(* IEC 61131-3 sources: 2026_Projet_YGO_ExcavatriceDragage/CODE_BACKUP/CODE_20260902_JoyAvantHoming_v0.6.27/G_CYCLE, 4 files *)

(* ---- FB_Cycle.st ---- *)
(* =======================================================================
   ⚙️ FB_Cycle — Séquenceur du cycle automatique (Grafcet de dragage)
   ───────────────────────────────────────────────────────────────
   🎯 Rôle : Automate de cycle automatique de dragage (X0 à X13 + STABILIZING)
   🔒 Sécurité : Gating par mode et homme-mort, repli STABILIZING sur défaut
   🔌 Interface : Demandes de mouvements (treuils, translation, benne)
   📄 Doc métier : DOC/AF/AF_Partie-04_Mode_SemiAuto_Sequenceur_v2.3.md
   ======================================================================= *)

FUNCTION_BLOCK PUBLIC FB_Cycle
VAR_INPUT
    // === COMMANDES & AUTORISATIONS ===
    Enable                  : BOOL;         // --> [CMD] Activation generale du sequenceur
    Reset                   : BOOL;         // --> [CMD] Acquittement defaut (front)
    PowerContactorEngaged   : BOOL;         // --> [SAFE] Chaine de securite OK
    EncoderFaultPresent     : BOOL;         // --> [SAFE] Defaut codeur agrege (cycle non autorise)
    Mode                    : E_Mode;       // --> [CMD] Mode arbitre (SEMI_AUTO pour instance cycle)
    JoystickDeflected       : BOOL;         // --> [CMD] Manche deflecte (non centre)
    DeadmanArmed            : BOOL;         // --> [CMD] Appui homme-mort (fenetre 3 s)
    HeartbeatIhmOk          : BOOL;         // --> [SAFE] IHM<->PLC valide

    // === COMMANDES OPERATEUR ===
    StartCycle              : BOOL;         // --> [CMD] Demande lancement / reprise (IHM)
    AbortCycle              : BOOL;         // --> [CMD] Demande abandon (IHM)

    // === CIBLES ET CONFIGURATION ===
    SelTarget               : INT;          // --> [CFG] Cible selectionnee (1=Tremie, 2=P2, 3=P1, 4=Maintenance)
    SetDepthM               : REAL;         // --> [CFG] Profondeur de consigne (negative)
    SetOffsetM              : REAL;         // --> [CFG] Ecart de fermeture benne cible

    // === FEEDBACKS CAPTEURS & MATERIEL ===
    KoboldContactFond       : BOOL;         // --> [HW] Retour dedie Kobold : TRUE = contact fond
    LimitLegalReached       : BOOL;         // --> [SAFE] Limite legale atteinte (descente interdite)
    LimitLegalDepthM        : REAL;         // --> [CFG] Profondeur legale minimale autorisee
    WinchSyncError          : BOOL;         // --> [SAFE] Desynchronisme bloquant M1/M2
    WinchSyncDeltaM         : REAL;         // --> [HW] Ecart codeurs M1/M2 pour diagnostic
    M1_CablePosM            : REAL;         // --> [HW] Position cable treuil M1 (recalee)
    M2_CablePosM            : REAL;         // --> [HW] Position cable treuil M2 (recalee)
    M1_MeasuredSpeedMps     : REAL;         // --> [HW] Vitesse lineaire mesuree M1 (m/s)
    M2_MeasuredSpeedMps     : REAL;         // --> [HW] Vitesse lineaire mesuree M2 (m/s)
    SpeedMismatchThresholdMps : REAL;       // --> [CFG] Seuil ecart vitesse ; 0 = controle desactive
    SpeedMismatchTimeout    : TIME;         // --> [CFG] Duree de confirmation ; 0 = controle desactive
    CableLimitM1AscentM     : REAL;         // --> [CFG] Limite haute d'exploitation M1

    // === FEEDBACKS TRANSLATION M3 ===
    Translation_At_P1           : BOOL;     // --> [HW] Capteur position P1 (arret travail)
    Translation_At_Tremie       : BOOL;     // --> [HW] Capteur fin de course tremie
    Translation_At_Maintenance : BOOL;     // --> [HW] Capteur fin de course maintenance
    Translation_Busy            : BOOL;     // --> [HW] Mouvement translation en cours
    Translation_Done            : BOOL;     // --> [HW] Cible translation atteinte

    // === FEEDBACKS BENNE ===
    Benne_Busy              : BOOL;         // --> [HW] Mouvement machoires benne en cours
    Benne_Done              : BOOL;         // --> [HW] Mouvement ouverture/fermeture termine
    Benne_IsOpen            : BOOL;         // --> [HW] Benne mecaniquement ouverte memorisee
    Benne_IsClosed          : BOOL;         // --> [HW] Benne mecaniquement fermee memorisee
    Benne_IsRoughlyClosed   : BOOL;         // --> [HW] Benne a peu pres fermee (tolerance matiere)

    // === REFERENCEMENT CODEURS ===
    HomedM1                 : BOOL;         // --> [HW] Codeur M1 reference
    HomedM2                 : BOOL;         // --> [HW] Codeur M2 reference
    TopPositionSensor       : BOOL;         // --> [HW] Capteur position haute (referencement)
    HomingRequest           : BOOL;         // --> [CMD] Demande de referencement (front)
END_VAR
VAR_OUTPUT
    // === ETATS IEC & DEFECTUOSITES ===
    Ready                   : BOOL;         // <-- [STAT] Sequenceur disponible
    Fault                   : ST_Fault;     // <-- [SAFE] Socle defaut transverse (live + latche)
    Lifecycle               : ST_Lifecycle; // <-- [STAT] Cycle de vie (Busy, Done, Waiting)
    SpeedMismatchMps        : REAL;         // <-- [DIAG] Ecart absolu vitesse M1/M2 (m/s)
    SpeedMismatchActive     : BOOL;         // <-- [DIAG] Seuil vitesse depasse sur cycle courant
    SpeedMismatchConfirmed  : BOOL;         // <-- [DIAG] Ecart vitesse confirme pendant timeout

    // === ORDRES ACTIONNEURS (COMMANDES STRUCTUREES) ===
    // Types de contrat inter-PRG uniques (ST_Program*Request) : FB_Cycle produit
    // directement les demandes consommées par PRG_04/05/07 — plus de DUT
    // ST_fbCycle_*CmdDemand redondants ni de re-mapping champ-à-champ (NC-090).
    WinchM1Cmd              : ST_ProgramWinchRequest;        // <-- [ACT] Demande treuil M1
    WinchM2Cmd              : ST_ProgramWinchRequest;        // <-- [ACT] Demande treuil M2
    TranslationCmd          : ST_ProgramTranslationRequest;  // <-- [ACT] Demande translation M3
    BucketCmd               : ST_ProgramBucketRequest;       // <-- [ACT] Demande benne

    // === METADONNEES & SYNOPTIQUE ===
    CycleStep               : E_CycleStep;          // <-- [STAT] Etape active du Grafcet
    CycleStateStr           : STRING(80);           // <-- [STAT] Libelle en clair de l'etape
    CycleStepAtError        : E_CycleStep;          // <-- [DIAG] Etape specifique au moment du defaut
    OperatorActionId        : WORD;                 // <-- [DIAG] ID action operateur requise
    OperatorAction          : STRING(120);          // <-- [DIAG] Message explicatif pour l'IHM
    ExpectedAxis            : E_OperatorAxis;       // <-- [STAT] Organe joystick/bouton attendu
    ExpectedDirection       : INT;                  // <-- [STAT] Sens attendu (-1, 0, +1)
    WaitingForOperator      : BOOL;                 // <-- [STAT] En attente d'une action operateur
    WaitingForProcess       : BOOL;                 // <-- [STAT] En attente d'une condition procede
    RequestActive           : BOOL;                 // <-- [STAT] Demande de mouvement active
END_VAR
VAR_IN_OUT
    // === STRUCTURES PARTAGEES & COMPTEURS ===
    SampleCount             : INT;          // <-> [BUS] Compteur de prelevements (RETAIN)
END_VAR
VAR
    // === DETECTEURS DE FRONTS ===
    ResetEdge               : R_TRIG;       // . [LOC] Detecteur front montant Reset
    StartEdge               : R_TRIG;       // . [LOC] Detecteur front montant StartCycle
    DeadmanArmedEdge        : R_TRIG;       // . [LOC] Detecteur front montant DeadmanArmed (demarrage joystick)
    AbortEdge               : R_TRIG;       // . [LOC] Detecteur front montant AbortCycle
    ErrorEdge               : R_TRIG;       // . [LOC] Detecteur front montant Error

    // === GATE CONTINU HOMME-MORT (permis par action hardware) ===
    ProcessPermitM1_Ascent   : BOOL; // . [LOC] Permis ascending treuil M1 = JoystickDeflected AND DeadmanArmed
    ProcessPermitM1_Descend  : BOOL; // . [LOC] Permis descending treuil M1 = JoystickDeflected AND DeadmanArmed
    ProcessPermitM2_Ascent   : BOOL; // . [LOC] Permis ascending treuil M2 = JoystickDeflected AND DeadmanArmed
    ProcessPermitM2_Descend  : BOOL; // . [LOC] Permis descending treuil M2 = JoystickDeflected AND DeadmanArmed
    ProcessPermitBucket_Open   : BOOL; // . [LOC] Permis ouverture benne = JoystickDeflected AND DeadmanArmed
    ProcessPermitBucket_Close   : BOOL; // . [LOC] Permis fermeture benne = JoystickDeflected AND DeadmanArmed
    ProcessPermitM3_Tremie          : BOOL; // . [LOC] Permis translation M3 cote tremie = JoystickDeflected AND DeadmanArmed
    ProcessPermitM3_Maintenance     : BOOL; // . [LOC] Permis translation M3 cote maintenance = JoystickDeflected AND DeadmanArmed

    // === COMPTEUR PRELEVEMENTS (garde de front) ===
    SampleCountDone         : BOOL := FALSE; // . [LOC] F2: front de comptage SampleCount (1 seul increment par cycle)

    // === ETATS INTERNES ===
    State                   : E_CycleStep := E_CycleStep.X0_PREPARATION; // . [LOC] Etape courante machine d'etat
    SavedState              : E_CycleStep := E_CycleStep.X0_PREPARATION; // . [LOC] Etape memorisee
    PausedState             : E_CycleStep := E_CycleStep.X0_PREPARATION; // . [LOC] Etape en pause lors de la bascule hors auto
    WaitingResume           : BOOL := FALSE;                             // . [LOC] En attente de validation consciente pour reprendre

    // === MEMORISATIONS & REGISTRES INTERNES ===
    TouchPositionM          : REAL;         // . [LOC] Position M1 memorisee lors du contact fond
    RaiseTargetM            : REAL;         // . [LOC] Profondeur de remontee memorisee
    SelectedWorkTarget      : INT;          // . [LOC] Cible de travail memorisee

    // === TEMPORISATEURS INTERNES ===
    DrainingTimer           : TON;          // . [LOC] Temporisateur de vidage (egouttage)
    StabilizationTimer      : TON;          // . [LOC] Temporisation maximale de remontee lente
    SpeedMismatchTimer      : TON;          // . [LOC] Confirmation temporelle ecart de vitesse
    StepMaxTimer            : TON;          // . [LOC] Tempo max d'etape

    // === CONSTANTES & CONFIGURATIONS INTERNES ===
    CtrlAscentDistM         : REAL := 2.0;      // . [LOC] Distance de remontee lente de controle
    CtrlAscentToleranceM    : REAL := 0.25;     // . [LOC] Ecart maximal admis entre codeurs
    CtrlAscentTimeout       : TIME := T#30s;    // . [LOC] Temps max pour zone de stabilisation
    DrainingTime            : TIME := T#5s;     // . [LOC] Temps d'egouttage par defaut
    StepMaxTimeout          : TIME := T#60s;    // . [LOC] Tempo max d'etape

    // === SOCLE DEFAUT TRANSVERSE ===
    instFault               : FB_FaultCore;                  // * [INST] Socle defaut transverse
    instCauses              : ARRAY[0..15] OF ST_FaultCause; // . [LOC] Table des causes de defaut
END_VAR

// === IMPLEMENTATION ===

{region "§1 Causes & Socle Défaut"}
// 🔑 1. FRONTS ET CAUSES
ResetEdge(CLK := Reset);
StartEdge(CLK := StartCycle);
DeadmanArmedEdge(CLK := DeadmanArmed);
AbortEdge(CLK := AbortCycle);

// ⏱️ Surveillance indépendante de la remontée lente
// X7_CTRL_ASCENT -> X8_ASCENT_LOADED : TON de stabilisation palier 1.
StabilizationTimer(IN := (State = E_CycleStep.X7_CTRL_ASCENT), PT := CtrlAscentTimeout);

// 📏 Comparaison vitesse réelle M1/M2
SpeedMismatchMps := ABS(M1_MeasuredSpeedMps - M2_MeasuredSpeedMps);
SpeedMismatchActive := (State = E_CycleStep.X7_CTRL_ASCENT)
                       AND JoystickDeflected
                       AND (SpeedMismatchThresholdMps > 0.0)
                       AND (SpeedMismatchTimeout > T#0ms)
                       AND (SpeedMismatchMps > SpeedMismatchThresholdMps);
// X7_CTRL_ASCENT -> STABILIZING : TON confirmation écart vitesse.
SpeedMismatchTimer(IN := SpeedMismatchActive, PT := SpeedMismatchTimeout);
SpeedMismatchConfirmed := SpeedMismatchTimer.Q;

// Tempo max d'étape (R5) — lancée SEULEMENT si pilotage joystick actif (pas de défaut au repos)
// Xi -> STABILIZING : TON backstop durée d'état pour tous les états de mouvement.
StepMaxTimer(IN := JoystickDeflected AND (State <> E_CycleStep.X0_PREPARATION)
                  AND (State <> E_CycleStep.X13_DONE_SYNC)
                  AND (State <> E_CycleStep.STABILIZING),
             PT := StepMaxTimeout);

// Table des causes de défaut
instCauses[0].Active   := LimitLegalReached AND (State = E_CycleStep.X4_DESCEND_OPEN);
instCauses[0].Latching := TRUE;
instCauses[0].Texte    := 'Limite legale de profondeur atteinte pendant descente';

instCauses[1].Active   := WinchSyncError AND (State <> E_CycleStep.X0_PREPARATION) AND (State <> E_CycleStep.STABILIZING);
instCauses[1].Latching := TRUE;
instCauses[1].Texte    := 'Desynchronisme treuils M1/M2 bloquant';

instCauses[2].Active   := SpeedMismatchConfirmed AND (State <> E_CycleStep.X0_PREPARATION) AND (State <> E_CycleStep.STABILIZING);
instCauses[2].Latching := TRUE;
instCauses[2].Texte    := 'Ecart de vitesse M1/M2 confirme en montee';

instCauses[3].Active   := NOT HeartbeatIhmOk AND (State <> E_CycleStep.X0_PREPARATION) AND (State <> E_CycleStep.STABILIZING);
instCauses[3].Latching := TRUE;
instCauses[3].Texte    := 'Perte communication IHM pendant cycle';

instCauses[4].Active   := StepMaxTimer.Q AND (State <> E_CycleStep.STABILIZING);
instCauses[4].Latching := TRUE;
instCauses[4].Texte    := 'Depassement tempo maximale d etape (blocage mouvement)';

instCauses[5].Active   := (StabilizationTimer.Q OR (ABS(M1_CablePosM - M2_CablePosM) > CtrlAscentToleranceM))
                          AND (State = E_CycleStep.X7_CTRL_ASCENT);
instCauses[5].Latching := TRUE;
instCauses[5].Texte    := 'Defaut de stabilisation / tolerance ecart codeurs en remontee controle';

// Appel du socle de défaut
instFault(Enable := Enable, Reset := Reset, Causes := instCauses);
Fault := instFault.Fault;
ErrorEdge(CLK := Fault.Error);
{endregion}

{region "§2 Gate securite & Bascule Mode"}
// 🛑 2. GATES DE SÉCURITÉ ET NEUTRALISATION
// Le mode SEMI_AUTO peut être sélectionné sous AU/défaut (FB_Modes), mais le cycle
// ne tourne JAMAIS sans puissance (PowerContactorEngaged) ni avec un codeur défaillant
// (EncoderFaultPresent) — les données de position invalides rendraient le Grafcet erroné.
IF NOT Enable OR NOT PowerContactorEngaged OR EncoderFaultPresent THEN
    WinchM1Cmd.RunRequest     := FALSE;
    WinchM1Cmd.ReqAscent      := FALSE;
    WinchM1Cmd.ReqDescend     := FALSE;
    WinchM1Cmd.StepTgt        := 0;

    WinchM2Cmd.RunRequest     := FALSE;
    WinchM2Cmd.ReqAscent      := FALSE;
    WinchM2Cmd.ReqDescend     := FALSE;
    WinchM2Cmd.StepTgt        := 0;

    TranslationCmd.ReqStart   := FALSE;
    TranslationCmd.PositionTgt  := 0;

    BucketCmd.ReqOpen         := FALSE;
    BucketCmd.ReqClose        := FALSE;
    BucketCmd.ReqKoboldMeasureEnable := FALSE;

    // Si on quitte le semi-auto alors qu'un cycle était en cours, on mémorise l'étape pour la pause
    IF (State <> E_CycleStep.X0_PREPARATION) AND (State <> E_CycleStep.X13_DONE_SYNC) AND (State <> E_CycleStep.STABILIZING) THEN
        PausedState := State;
        WaitingResume := TRUE;
    END_IF;

    CycleStep            := State;
    CycleStateStr        := 'Cycle desactive : securite/codeur/mode';
    Ready                := FALSE;
    Lifecycle.Busy       := FALSE;
    Lifecycle.Done       := FALSE;
    SpeedMismatchTimer(IN := FALSE, PT := SpeedMismatchTimeout);
    SpeedMismatchMps := 0.0;
    SpeedMismatchActive := FALSE;
    SpeedMismatchConfirmed := FALSE;
    OperatorActionId := 0;
    IF EncoderFaultPresent THEN
        OperatorAction := 'Cycle non autorise : defaut codeur present. Reinitialiser le defaut codeur.';
    ELSE
        OperatorAction := 'Passer en mode Semi-Auto et engager la securite pour activer le cycle.';
    END_IF;
    ExpectedAxis := E_OperatorAxis.NONE;
    ExpectedDirection := 0;
    WaitingForOperator := FALSE;
    WaitingForProcess := FALSE;
    RequestActive := FALSE;
    RETURN;
END_IF;

Ready := Enable AND NOT Fault.Latched;

// 🛡️ Gate continu homme-mort : le mouvement n'est autorisé que si le manche est
// défléchi (JoystickDeflected) ET l'homme-mort est armé (DeadmanArmed). Chaque
// commande de mouvement est gatée par ce permis à chaque scan (pas seulement au
// démarrage). Le séquenceur (transitions X0→X13) reste piloté par JoystickDeflected.
ProcessPermitM1_Ascent        := JoystickDeflected AND DeadmanArmed;
ProcessPermitM1_Descend      := JoystickDeflected AND DeadmanArmed;
ProcessPermitM2_Ascent        := JoystickDeflected AND DeadmanArmed;
ProcessPermitM2_Descend      := JoystickDeflected AND DeadmanArmed;
ProcessPermitBucket_Open := JoystickDeflected AND DeadmanArmed;
ProcessPermitBucket_Close := JoystickDeflected AND DeadmanArmed;
ProcessPermitM3_Tremie        := JoystickDeflected AND DeadmanArmed;
ProcessPermitM3_Maintenance   := JoystickDeflected AND DeadmanArmed;

// Au retour en Semi-Auto, si une étape était en cours, on exige une reprise consciente
IF WaitingResume THEN
    // 🔒 Sécurité anti-redémarrage automatique (AF-04 §4.1) : le cycle ne reprend
    // PAS sur manche + homme-mort seuls. Il reste en attente d'un geste conscient
    // (StartCycle) avant de restaurer l'étape mémorisée.
    IF StartEdge.Q THEN
        State := PausedState;   // reprise consciente : restaure l'étape mémorisée
        WaitingResume := FALSE;
    ELSE
        // Hold : neutralise toute demande de mouvement et affiche l'attente.
        WinchM1Cmd.RunRequest := FALSE; WinchM1Cmd.ReqAscent := FALSE; WinchM1Cmd.ReqDescend := FALSE; WinchM1Cmd.StepTgt := 0;
        WinchM2Cmd.RunRequest := FALSE; WinchM2Cmd.ReqAscent := FALSE; WinchM2Cmd.ReqDescend := FALSE; WinchM2Cmd.StepTgt := 0;
        TranslationCmd.ReqStart := FALSE; TranslationCmd.PositionTgt := 0;
        BucketCmd.ReqOpen := FALSE; BucketCmd.ReqClose := FALSE; BucketCmd.ReqKoboldMeasureEnable := FALSE;
        CycleStep := PausedState;
        CycleStateStr := 'Cycle en pause : reprise consciente requise (StartCycle)';
        Lifecycle.Busy := FALSE;
        Lifecycle.Done := FALSE;
        ExpectedAxis := E_OperatorAxis.BUTTON;
        ExpectedDirection := 0;
        WaitingForOperator := TRUE;
        WaitingForProcess := FALSE;
        OperatorActionId := 16#0400;
        OperatorAction := 'Reprendre le cycle : appuyer sur StartCycle (geste conscient).';
        RequestActive := FALSE;
    END_IF;
END_IF;

// 🧊 R9 — capture l'étape spécifique AVANT la bascule vers STABILIZING
IF ErrorEdge.Q THEN
    CycleStepAtError := State;
    State := E_CycleStep.STABILIZING;
    WaitingResume := FALSE;   // un défaut abroge la reprise consciente : repli STABILIZING
END_IF;

IF ResetEdge.Q THEN
    SavedState := E_CycleStep.X0_PREPARATION;
    IF State = E_CycleStep.STABILIZING THEN
        State := E_CycleStep.X0_PREPARATION;
    END_IF;
END_IF;

// Gestion de l'Abandon explicite
IF AbortEdge.Q THEN
    State := E_CycleStep.X0_PREPARATION;
    WaitingResume := FALSE;
    PausedState := E_CycleStep.X0_PREPARATION;
END_IF;

// SEMI_AUTO : FB_Cycle est le SEUL producteur des demandes benne. Les champs
// assistants (DiveSearch/ExtractionAssist) sont inactifs en cycle automatique
// -> valeurs neutres déterministes (identiques à la branche SEMI_AUTO de PRG_03).
BucketCmd.DescendPermitDiveBucketOpen := TRUE;
BucketCmd.ExtractionControlActive := FALSE;
BucketCmd.MinStepDown := 0;
{endregion}

{region "§3 Machine etat cycle automatique"}
// 🔁 2. LOGIQUE DU SÉQUENCEUR (Machine d'état) — CASE sur enum unique (R1)
// Pendant une reprise consciente (WaitingResume), le séquenceur est gelé :
// l'étape mémorisée ne s'exécute pas tant que StartCycle n'a pas été appuyé.
IF NOT WaitingResume THEN
CASE State OF

    E_CycleStep.X0_PREPARATION:
        CycleStep := E_CycleStep.X0_PREPARATION;
        CycleStateStr := 'X0 - Verification coherence systeme';
        WinchM1Cmd.RunRequest := FALSE; WinchM1Cmd.ReqAscent := FALSE; WinchM1Cmd.ReqDescend := FALSE; WinchM1Cmd.StepTgt := 0;
        WinchM2Cmd.RunRequest := FALSE; WinchM2Cmd.ReqAscent := FALSE; WinchM2Cmd.ReqDescend := FALSE; WinchM2Cmd.StepTgt := 0;
        TranslationCmd.ReqStart := FALSE; TranslationCmd.PositionTgt := 0;
        BucketCmd.ReqOpen := FALSE; BucketCmd.ReqClose := FALSE; BucketCmd.ReqKoboldMeasureEnable := FALSE;
        Lifecycle.Busy := FALSE;
        Lifecycle.Done := FALSE;
        ExpectedAxis := E_OperatorAxis.BUTTON;
        ExpectedDirection := 0;
        WaitingForOperator := TRUE;
        WaitingForProcess := FALSE;
        OperatorActionId := 16#0400;
        OperatorAction := 'Demander le demarrage du cycle (Bouton IHM ou armement Homme-Mort).';
        SampleCountDone := FALSE;   // F2: réarmement du front de comptage à chaque entrée en X0

        // Transition si système sain et réarmé (front reset ou démarrage).
        // 🔫 D2 : démarrage par bouton IHM (StartEdge) OU armement homme-mort joystick
        IF (StartEdge.Q OR DeadmanArmedEdge.Q) AND NOT Fault.Latched THEN
            WaitingResume := FALSE;
            State := E_CycleStep.X1_HOMING;
        END_IF;

    E_CycleStep.X1_HOMING:
        CycleStep := E_CycleStep.X1_HOMING;
        CycleStateStr := 'X1 - Referencement codeurs (vitesses lentes)';
        Lifecycle.Busy := TRUE;
        Lifecycle.Done := FALSE;
        ExpectedAxis := E_OperatorAxis.JOYSTICK_Y;
        ExpectedDirection := 1;
        WaitingForOperator := NOT JoystickDeflected;
        WaitingForProcess := JoystickDeflected;
        OperatorActionId := 16#0401;
        OperatorAction := 'Maintenir la montee lente vers les capteurs de referencement.';

        // Vitesses lentes pour chercher capteur top + référencement
        IF NOT HomedM1 OR NOT HomedM2 THEN
            WinchM1Cmd.RunRequest := ProcessPermitM1_Ascent;
            WinchM1Cmd.ReqAscent := TRUE; WinchM1Cmd.ReqDescend := FALSE;   // montée lente vers capteur top
            WinchM1Cmd.StepTgt := 1;
            WinchM2Cmd.RunRequest := ProcessPermitM2_Ascent;
            WinchM2Cmd.ReqAscent := TRUE; WinchM2Cmd.ReqDescend := FALSE;
            WinchM2Cmd.StepTgt := 1;
            IF HomingRequest THEN
                State := E_CycleStep.X2_WORK_POS_SELECT;
            END_IF;
        ELSE
            // déjà homé → passe vite
            State := E_CycleStep.X2_WORK_POS_SELECT;
        END_IF;

    E_CycleStep.X2_WORK_POS_SELECT:
        CycleStep := E_CycleStep.X2_WORK_POS_SELECT;
        CycleStateStr := 'X2 - Selection position travail';
        Lifecycle.Busy := TRUE;
        Lifecycle.Done := FALSE;
        ExpectedAxis := E_OperatorAxis.JOYSTICK_X;
        ExpectedDirection := 0;
        WaitingForOperator := (SelTarget = 0) OR NOT JoystickDeflected;
        WaitingForProcess := (SelTarget <> 0) AND JoystickDeflected;
        OperatorActionId := 16#0402;
        OperatorAction := 'Selectionner la cible et maintenir la translation vers la position de travail.';

        IF (SelTarget = 1) OR (SelTarget = 3) OR (SelTarget = 4) THEN
            SelectedWorkTarget := SelTarget;
            TranslationCmd.PositionTgt := SelTarget;
            TranslationCmd.ReqStart := ProcessPermitM3_Tremie;
            // Arrivée à la cible (Trémie/P1/Maintenance)
            IF JoystickDeflected AND (
                (SelTarget = 1 AND Translation_At_Tremie) OR
                (SelTarget = 3 AND Translation_At_P1) OR
                (SelTarget = 4 AND Translation_At_Maintenance)) THEN
                TranslationCmd.ReqStart := FALSE;
                State := E_CycleStep.X3_OPEN_BUCKET;
            END_IF;
        END_IF;

    E_CycleStep.X3_OPEN_BUCKET:
        CycleStep := E_CycleStep.X3_OPEN_BUCKET;
        CycleStateStr := 'X3 - Ouverture benne';
        Lifecycle.Busy := TRUE;
        Lifecycle.Done := FALSE;
        ExpectedAxis := E_OperatorAxis.JOYSTICK_Y;
        ExpectedDirection := 0;
        WaitingForOperator := NOT JoystickDeflected;
        WaitingForProcess := JoystickDeflected;
        OperatorActionId := 16#0403;
        OperatorAction := 'Maintenir le joystick : ouverture complete de la benne.';

        IF Benne_IsOpen THEN
            State := E_CycleStep.X4_DESCEND_OPEN;
        ELSE
            BucketCmd.ReqOpen := ProcessPermitBucket_Open;
            IF JoystickDeflected AND Benne_Done AND Benne_IsOpen THEN
                BucketCmd.ReqOpen := FALSE;
                State := E_CycleStep.X4_DESCEND_OPEN;
            END_IF;
        END_IF;

    E_CycleStep.X4_DESCEND_OPEN:
        CycleStep := E_CycleStep.X4_DESCEND_OPEN;
        CycleStateStr := 'X4 - Plongee benne ouverte (synchro)';
        Lifecycle.Busy := TRUE;
        Lifecycle.Done := FALSE;
        ExpectedAxis := E_OperatorAxis.JOYSTICK_Y;
        ExpectedDirection := -1;
        WaitingForOperator := NOT JoystickDeflected;
        WaitingForProcess := JoystickDeflected;
        OperatorActionId := 16#0404;
        OperatorAction := 'Maintenir la descente : plongee synchro et detection fond Kobold.';

        // M1 et M2 descendent ensemble (synchro gérée en aval)
        WinchM1Cmd.RunRequest := ProcessPermitM1_Descend;
        WinchM1Cmd.ReqAscent := FALSE; WinchM1Cmd.ReqDescend := TRUE;
        WinchM1Cmd.StepTgt  := 3;
        WinchM2Cmd.RunRequest := ProcessPermitM2_Descend;
        WinchM2Cmd.ReqAscent := FALSE; WinchM2Cmd.ReqDescend := TRUE;
        WinchM2Cmd.StepTgt  := 3;
        BucketCmd.ReqKoboldMeasureEnable := ProcessPermitM1_Descend;

        // Transition uniquement sur le retour dédié Kobold.
        IF JoystickDeflected AND KoboldContactFond THEN
            WinchM1Cmd.RunRequest := FALSE;
            WinchM2Cmd.RunRequest := FALSE;
            BucketCmd.ReqKoboldMeasureEnable := FALSE;
            TouchPositionM := M1_CablePosM;
            IF LimitLegalDepthM < -0.01 THEN
                RaiseTargetM := MAX(TouchPositionM + 0.5, LimitLegalDepthM + 0.5);
            ELSE
                RaiseTargetM := TouchPositionM + 0.5;
            END_IF;
            State := E_CycleStep.X5_BOTTOM_CONFIRMED;
        END_IF;

    E_CycleStep.X5_BOTTOM_CONFIRMED:
        CycleStep := E_CycleStep.X5_BOTTOM_CONFIRMED;
        CycleStateStr := 'X5 - Fond confirme : remontee securisee';
        Lifecycle.Busy := TRUE;
        Lifecycle.Done := FALSE;
        ExpectedAxis := E_OperatorAxis.JOYSTICK_Y;
        ExpectedDirection := 1;
        WaitingForOperator := NOT JoystickDeflected;
        WaitingForProcess := JoystickDeflected;
        OperatorActionId := 16#0405;
        OperatorAction := 'Fond confirme : maintenir la montee jusqu a la hauteur de fermeture.';

        WinchM1Cmd.RunRequest := ProcessPermitM1_Ascent;
        WinchM1Cmd.ReqAscent := TRUE; WinchM1Cmd.ReqDescend := FALSE;
        WinchM1Cmd.StepTgt := 1;
        WinchM2Cmd.RunRequest := ProcessPermitM2_Ascent;
        WinchM2Cmd.ReqAscent := TRUE; WinchM2Cmd.ReqDescend := FALSE;
        WinchM2Cmd.StepTgt := 1;

        IF JoystickDeflected AND (M1_CablePosM >= RaiseTargetM) AND (M2_CablePosM >= RaiseTargetM) THEN
            WinchM1Cmd.RunRequest := FALSE;
            WinchM2Cmd.RunRequest := FALSE;
            State := E_CycleStep.X6_CLOSE_BUCKET;
        END_IF;

    E_CycleStep.X6_CLOSE_BUCKET:
        CycleStep := E_CycleStep.X6_CLOSE_BUCKET;
        CycleStateStr := 'X6 - Fermeture benne (tolerance a peu pres ferme)';
        Lifecycle.Busy := TRUE;
        Lifecycle.Done := FALSE;
        ExpectedAxis := E_OperatorAxis.JOYSTICK_Y;
        ExpectedDirection := 1;
        WaitingForOperator := NOT JoystickDeflected;
        WaitingForProcess := JoystickDeflected;
        OperatorActionId := 16#0406;
        OperatorAction := 'Maintenir la commande : fermeture de la benne.';

        WinchM1Cmd.RunRequest := FALSE;
        // L'ordre benne reste soumis au même homme-mort que le cycle : aucune
        // commande d'actionneur ne doit survivre à la perte du permis opérateur.
        BucketCmd.ReqClose := ProcessPermitBucket_Close;

        IF JoystickDeflected AND (Benne_Done AND (Benne_IsClosed OR Benne_IsRoughlyClosed)) THEN
            BucketCmd.ReqClose := FALSE;
            State := E_CycleStep.X7_CTRL_ASCENT;
        END_IF;

    E_CycleStep.X7_CTRL_ASCENT:
        CycleStep := E_CycleStep.X7_CTRL_ASCENT;
        CycleStateStr := 'X7 - Remontee lente de controle';
        Lifecycle.Busy := TRUE;
        Lifecycle.Done := FALSE;
        ExpectedAxis := E_OperatorAxis.JOYSTICK_Y;
        ExpectedDirection := 1;
        WaitingForOperator := NOT JoystickDeflected;
        WaitingForProcess := JoystickDeflected;
        OperatorActionId := 16#0407;
        OperatorAction := 'Maintenir la montee lente : palier de controle et synchronisme.';

        WinchM1Cmd.RunRequest := ProcessPermitM1_Ascent;
        WinchM1Cmd.ReqAscent := TRUE; WinchM1Cmd.ReqDescend := FALSE;
        WinchM1Cmd.StepTgt  := 1;
        WinchM2Cmd.RunRequest := ProcessPermitM2_Ascent;
        WinchM2Cmd.ReqAscent := TRUE; WinchM2Cmd.ReqDescend := FALSE;
        WinchM2Cmd.StepTgt  := 1;

        IF JoystickDeflected
           AND (M1_CablePosM >= (TouchPositionM + CtrlAscentDistM))
           AND (M2_CablePosM >= (TouchPositionM + CtrlAscentDistM))
           AND (ABS(M1_CablePosM - M2_CablePosM) <= CtrlAscentToleranceM) THEN
            State := E_CycleStep.X8_ASCENT_LOADED;
        END_IF;

    E_CycleStep.X8_ASCENT_LOADED:
        CycleStep := E_CycleStep.X8_ASCENT_LOADED;
        CycleStateStr := 'X8 - Remontee en charge';
        Lifecycle.Busy := TRUE;
        Lifecycle.Done := FALSE;
        ExpectedAxis := E_OperatorAxis.JOYSTICK_Y;
        ExpectedDirection := 1;
        WaitingForOperator := NOT JoystickDeflected;
        WaitingForProcess := JoystickDeflected;
        OperatorActionId := 16#0408;
        OperatorAction := 'Maintenir la montee en charge jusqu a la limite haute.';

        WinchM1Cmd.RunRequest := ProcessPermitM1_Ascent;
        WinchM1Cmd.ReqAscent := TRUE; WinchM1Cmd.ReqDescend := FALSE;
        WinchM1Cmd.StepTgt  := 4;
        WinchM2Cmd.RunRequest := ProcessPermitM2_Ascent;
        WinchM2Cmd.ReqAscent := TRUE; WinchM2Cmd.ReqDescend := FALSE;
        WinchM2Cmd.StepTgt  := 4;

        IF JoystickDeflected AND M1_CablePosM >= CableLimitM1AscentM THEN
            WinchM1Cmd.RunRequest := FALSE;
            WinchM2Cmd.RunRequest := FALSE;
            State := E_CycleStep.X9_DRAIN_PAUSE;
        END_IF;

    E_CycleStep.X9_DRAIN_PAUSE:
        CycleStep := E_CycleStep.X9_DRAIN_PAUSE;
        CycleStateStr := 'X9 - Egouttage du godet en cours';
        Lifecycle.Busy := TRUE;
        Lifecycle.Done := FALSE;
        ExpectedAxis := E_OperatorAxis.NONE;
        ExpectedDirection := 0;
        WaitingForOperator := FALSE;
        WaitingForProcess := TRUE;
        OperatorActionId := 16#0409;
        OperatorAction := 'Egouttage du godet en cours (temporisation).';
        WinchM1Cmd.RunRequest := FALSE;
        WinchM2Cmd.RunRequest := FALSE;

        DrainingTimer(IN := TRUE, PT := DrainingTime);
        IF JoystickDeflected AND DrainingTimer.Q THEN
            DrainingTimer(IN := FALSE);
            State := E_CycleStep.X10_TRANSLATE_DUMP;
        END_IF;

    E_CycleStep.X10_TRANSLATE_DUMP:
        CycleStep := E_CycleStep.X10_TRANSLATE_DUMP;
        CycleStateStr := 'X10 - Deplacement vers tremie (grille/crible libres)';
        Lifecycle.Busy := TRUE;
        Lifecycle.Done := FALSE;
        ExpectedAxis := E_OperatorAxis.JOYSTICK_X;
        ExpectedDirection := -1;
        WaitingForOperator := NOT JoystickDeflected;
        WaitingForProcess := JoystickDeflected;
        OperatorActionId := 16#040A;
        OperatorAction := 'Maintenir la translation vers la tremie de dechargement.';

        TranslationCmd.PositionTgt := 1; // Trémie
        TranslationCmd.ReqStart := ProcessPermitM3_Tremie;

        IF JoystickDeflected AND Translation_At_Tremie THEN
            TranslationCmd.ReqStart := FALSE;
            State := E_CycleStep.X11_OPEN_DUMP;
        END_IF;

    E_CycleStep.X11_OPEN_DUMP:
        CycleStep := E_CycleStep.X11_OPEN_DUMP;
        CycleStateStr := 'X11 - Vidange / ouverture du godet (montee possible, descente ouvre)';
        Lifecycle.Busy := TRUE;
        Lifecycle.Done := FALSE;
        ExpectedAxis := E_OperatorAxis.JOYSTICK_Y;
        ExpectedDirection := -1;
        WaitingForOperator := NOT JoystickDeflected;
        WaitingForProcess := JoystickDeflected;
        OperatorActionId := 16#040B;
        OperatorAction := 'Deflechir vers le bas pour ouvrir la benne et vider la charge.';

        // X11 est une ouverture par déflexion vers le bas : la direction doit
        // être écrite avant d'être évaluée (ne jamais tester la valeur du scan
        // précédent). Les deux treuils restent synchrones et sous homme-mort.
        WinchM1Cmd.ReqAscent := FALSE; WinchM1Cmd.ReqDescend := TRUE;
        WinchM1Cmd.RunRequest := ProcessPermitM1_Descend;
        WinchM1Cmd.StepTgt  := 1;
        WinchM2Cmd.ReqAscent := FALSE; WinchM2Cmd.ReqDescend := TRUE;
        WinchM2Cmd.RunRequest := ProcessPermitM2_Descend;
        WinchM2Cmd.StepTgt  := 1;

        BucketCmd.ReqOpen := ProcessPermitBucket_Open AND WinchM1Cmd.ReqDescend;

        IF JoystickDeflected AND Benne_Done AND Benne_IsOpen THEN
            BucketCmd.ReqOpen := FALSE;
            State := E_CycleStep.X13_DONE_SYNC;
        END_IF;

    E_CycleStep.X13_DONE_SYNC:
        CycleStep := E_CycleStep.X13_DONE_SYNC;
        CycleStateStr := 'X13 - Cycle automatique complete - pret';
        WinchM1Cmd.RunRequest := FALSE;
        WinchM2Cmd.RunRequest := FALSE;
        TranslationCmd.ReqStart := FALSE;
        Lifecycle.Done := TRUE;
        Lifecycle.Busy := FALSE;
        ExpectedAxis := E_OperatorAxis.BUTTON;
        ExpectedDirection := 0;
        WaitingForOperator := TRUE;
        WaitingForProcess := FALSE;
        OperatorActionId := 16#040D;
        OperatorAction := 'Cycle termine avec succes. Relancer un nouveau cycle.';

        // Compteur de prélèvements (RETAIN) — F2: incrément cadré par front (1 seul par cycle)
        IF NOT SampleCountDone THEN
            SampleCount := SampleCount + 1;
            SampleCountDone := TRUE;
        END_IF;

        IF StartEdge.Q THEN
            SampleCountDone := FALSE;
            Lifecycle.Done := FALSE;
            State := E_CycleStep.X0_PREPARATION;
        END_IF;

    E_CycleStep.STABILIZING:
        CycleStep := E_CycleStep.STABILIZING;
        CycleStateStr := 'X14 - Cycle en attente / stabilisation (STAB)';
        WinchM1Cmd.RunRequest := FALSE; WinchM1Cmd.ReqAscent := FALSE; WinchM1Cmd.ReqDescend := FALSE;
        WinchM2Cmd.RunRequest := FALSE; WinchM2Cmd.ReqAscent := FALSE; WinchM2Cmd.ReqDescend := FALSE;
        TranslationCmd.ReqStart := FALSE;
        BucketCmd.ReqOpen := FALSE;
        BucketCmd.ReqClose := FALSE;
        BucketCmd.ReqKoboldMeasureEnable := FALSE;   // Coupure contacteur Kobold au repli defaut (0 ordre residuel)
        Lifecycle.Busy := FALSE;
        Lifecycle.Done := FALSE;
        ExpectedAxis := E_OperatorAxis.BUTTON;
        ExpectedDirection := 0;
        WaitingForOperator := TRUE;
        WaitingForProcess := FALSE;
        OperatorActionId := 16#0480;
        OperatorAction := 'Cycle stabilise sur anomalie : acquitter le defaut pour reinitialiser.';

END_CASE;
END_IF;
{endregion}

{region "§4 Repli homme mort & Syntheses"}
// 🛑 Relâchement du manche (retour au centre) OU de l'homme-mort : neutralisation
// des demandes actives. Gate continu : aucune commande d'actionneur ne survit à la
// perte du permis opérateur (manche défléchi ET homme-mort armé).
IF Lifecycle.Busy AND NOT ProcessPermitM1_Ascent THEN
    WinchM1Cmd.RunRequest := FALSE;
    WinchM2Cmd.RunRequest := FALSE;
    TranslationCmd.ReqStart := FALSE;
    BucketCmd.ReqOpen := FALSE;
    BucketCmd.ReqClose := FALSE;
    BucketCmd.ReqKoboldMeasureEnable := FALSE;
END_IF;

RequestActive := WinchM1Cmd.RunRequest OR WinchM2Cmd.RunRequest OR TranslationCmd.ReqStart OR BucketCmd.ReqOpen OR BucketCmd.ReqClose OR BucketCmd.ReqKoboldMeasureEnable; // Somme logique complete des demandes (contacteur Kobold inclus)
{endregion}

END_FUNCTION_BLOCK

(* ---- FB_DiveSearch.st ---- *)
(* =======================================================================
   FB_DiveSearch - Assistance plongee et recherche du fond Kobold
   Role : qualifier l'immersion et autoriser la descente assistee.
   Interface : contrat standard + bus Inputs/Outputs.
   Documentation : DOC/AF/AF_Partie-04_Mode_SemiAuto_Sequenceur_v2.3.md
   ======================================================================= *)
FUNCTION_BLOCK FB_DiveSearch
VAR_INPUT
    // === CONTRAT STANDARD ===
    Enable                  : BOOL;                   // --> [CMD] Autorisation generale du FB
    Reset                   : BOOL;                   // --> [CMD] Acquittement defaut sur front

    // === BUS FONCTIONNEL ===
    Inputs                  : ST_fbDiveSearch_Inputs; // --> [BUS] Commande, capteurs et reglages
END_VAR
VAR_OUTPUT
    // === STATUT IEC ===
    Ready                   : BOOL;                   // <-- [STAT] FB pret a fonctionner
    Fault                   : ST_Fault;               // <-- [DIAG] Defaut live et latche
    Lifecycle               : ST_Lifecycle;           // <-- [STAT] Cycle en cours / termine

    // === BUS FONCTIONNEL ===
    Outputs                 : ST_fbDiveSearch_Outputs;// <-- [BUS] Etat, permis et diagnostic
END_VAR
VAR
    // === SOUS-INSTANCES & FRONTS ===
    ResetEdge               : R_TRIG;                 // . [LOC] Front Reset
    ErrorEdge               : R_TRIG;                 // . [LOC] Apparition d'un defaut
    KoboldRiseEdge          : R_TRIG;                 // . [LOC] Entree dans l'eau
    KoboldFallEdge          : F_TRIG;                 // . [LOC] Sortie de l'eau / fond
    instFault               : FB_FaultCore;           // * [INST] Socle defaut transverse
    instCauses              : ARRAY[0..15] OF ST_FaultCause; // . [LOC] Causes nommees

    // === CALCULS DE GARDE ===
    ImmersionCourse_M          : REAL;                // . [LOC] Course maximale vers immersion (m)
    BottomCourse_M             : REAL;                // . [LOC] Course maximale vers fond (m)
    CalculatedImmersionTimeout : TIME;                // . [LOC] Timeout immersion calcule
    CalculatedBottomTimeout    : TIME;                // . [LOC] Timeout fond calcule
    EffectiveDiveSpeedMin_Mps  : REAL;                // . [LOC] Vitesse minimale appliquee (m/s)
    EffectiveTimeoutMargin     : REAL;                // . [LOC] Marge appliquee au calcul
    EffectiveTimeoutMinCourse_M: REAL;                // . [LOC] Plancher de course applique (m)
    EffectiveTimeoutMaxCourse_M: REAL;                // . [LOC] Plafond de course applique (m)
    EffectiveSecToMs            : REAL;               // . [LOC] Conversion secondes/millisecondes

    // === MEMORISATIONS & TEMPORISATIONS ===
    ImmersionTimerAcc       : TIME := T#0ms;          // . [LOC] Temps effectif de recherche immersion
    BottomTimerAcc          : TIME := T#0ms;          // . [LOC] Temps effectif de recherche fond
    PrevState               : E_DiveSearchState;      // . [LOC] Etat du scan precedent
    ImmersionConfirmed      : BOOL;                   // . [LOC] Immersion validee
    StepAtFaultCaptured     : BOOL;                   // . [LOC] Etape de defaut deja figee

    // === CAUSES INTERNES ===
    ErrorCausePresent       : BOOL;                   // . [LOC] Parametrage invalide
    SeqErrorFault           : BOOL;                   // . [LOC] Incoherence de sequence
    Palier5ForbiddenFault   : BOOL;                   // . [LOC] Palier 5 interdit sous Kobold
    TimeoutImmersionFault   : BOOL;                   // . [LOC] Timeout recherche immersion
    TimeoutBottomFault      : BOOL;                   // . [LOC] Timeout recherche fond
    DescentActive           : BOOL;                   // . [LOC] Descending demandee et autorisee
END_VAR

{region "§1 Fronts, calculs et causes"}
ResetEdge(CLK := Reset);
KoboldRiseEdge(CLK := Inputs.KoboldImmersed);
KoboldFallEdge(CLK := Inputs.KoboldImmersed);

// Les valeurs par defaut du DUT couvrent l'appel sans configuration explicite.
// Le repli runtime protege aussi un appel avec une structure entierement nulle.
EffectiveDiveSpeedMin_Mps := Inputs.Config.DiveSpeedMin_Mps;
IF EffectiveDiveSpeedMin_Mps <= 0.0 THEN EffectiveDiveSpeedMin_Mps := 0.15; END_IF;
EffectiveTimeoutMargin := Inputs.Config.TimeoutMarginFactor;
IF EffectiveTimeoutMargin <= 0.0 THEN EffectiveTimeoutMargin := 1.5; END_IF;
EffectiveTimeoutMinCourse_M := Inputs.Config.TimeoutMinCourse_M;
IF EffectiveTimeoutMinCourse_M <= 0.0 THEN EffectiveTimeoutMinCourse_M := 1.0; END_IF;
EffectiveTimeoutMaxCourse_M := Inputs.Config.TimeoutMaxCourse_M;
IF EffectiveTimeoutMaxCourse_M < EffectiveTimeoutMinCourse_M THEN EffectiveTimeoutMaxCourse_M := 200.0; END_IF;
EffectiveSecToMs := Inputs.Config.SecToMs;
IF EffectiveSecToMs <= 0.0 THEN EffectiveSecToMs := 1000.0; END_IF;

ErrorCausePresent := (Inputs.CycleTime <= T#0ms)
                 OR (NOT Inputs.BypassPreconditions AND (
                       (Inputs.DiveStartMin_M < Inputs.ImmersionUpper_M)
                    OR (Inputs.ImmersionUpper_M <= Inputs.ImmersionLower_M)
                    OR (Inputs.ImmersionLower_M <= Inputs.LimitLegalDepthMin_M)
                    OR (Inputs.CableLimitAscent_M <= Inputs.ImmersionLower_M)));

ImmersionCourse_M := LIMIT(EffectiveTimeoutMinCourse_M,
                           Inputs.CableLimitAscent_M - Inputs.ImmersionLower_M,
                           EffectiveTimeoutMaxCourse_M);
BottomCourse_M := LIMIT(EffectiveTimeoutMinCourse_M,
                        Inputs.ImmersionLower_M - Inputs.LimitLegalDepthMin_M,
                        EffectiveTimeoutMaxCourse_M);
CalculatedImmersionTimeout := UDINT_TO_TIME(REAL_TO_UDINT(
    ImmersionCourse_M / EffectiveDiveSpeedMin_Mps * EffectiveTimeoutMargin * EffectiveSecToMs));
CalculatedBottomTimeout := UDINT_TO_TIME(REAL_TO_UDINT(
    BottomCourse_M / EffectiveDiveSpeedMin_Mps * EffectiveTimeoutMargin * EffectiveSecToMs));

IF (Outputs.StepState = E_DiveSearchState.SEARCHING_IMMERSION)
   AND Inputs.MotionRequestActive AND (Inputs.MotionDirection = -1) THEN
    ImmersionTimerAcc := ImmersionTimerAcc + Inputs.CycleTime;
    IF ImmersionTimerAcc >= CalculatedImmersionTimeout THEN TimeoutImmersionFault := TRUE; END_IF;
END_IF;

IF (Outputs.StepState = E_DiveSearchState.SEARCHING_BOTTOM)
   AND Inputs.MotionRequestActive AND (Inputs.MotionDirection = -1) THEN
    BottomTimerAcc := BottomTimerAcc + Inputs.CycleTime;
    IF BottomTimerAcc >= CalculatedBottomTimeout THEN TimeoutBottomFault := TRUE; END_IF;
END_IF;

IF ResetEdge.Q AND NOT ErrorCausePresent AND NOT Inputs.KoboldImmersed
   AND NOT Inputs.MotionRequestActive AND NOT (Inputs.CurrentSpeedStep > 4) THEN
    SeqErrorFault := FALSE;
    Palier5ForbiddenFault := FALSE;
    TimeoutImmersionFault := FALSE;
    TimeoutBottomFault := FALSE;
    ImmersionTimerAcc := T#0ms;
    BottomTimerAcc := T#0ms;
    ImmersionConfirmed := FALSE;
    Outputs.BottomTouchConfirmed := FALSE;
    Outputs.StepAtFault := E_DiveSearchState.WAIT_PRECONDITIONS;
    StepAtFaultCaptured := FALSE;
    Outputs.StepState := E_DiveSearchState.WAIT_PRECONDITIONS;
END_IF;

instCauses[0].Active := SeqErrorFault;
instCauses[0].Latching := TRUE;
instCauses[0].Texte := 'Incoherence sequence immersion Kobold';
instCauses[1].Active := ErrorCausePresent;
instCauses[1].Latching := TRUE;
instCauses[1].Texte := 'Parametrage invalide des seuils de plongee';
instCauses[2].Active := Palier5ForbiddenFault;
instCauses[2].Latching := TRUE;
instCauses[2].Texte := 'Palier 5 interdit pendant la mesure Kobold';
instCauses[3].Active := TimeoutImmersionFault;
instCauses[3].Latching := TRUE;
instCauses[3].Texte := 'Timeout recherche immersion Kobold';
instCauses[4].Active := TimeoutBottomFault;
instCauses[4].Latching := TRUE;
instCauses[4].Texte := 'Timeout recherche fond Kobold';

instFault(Enable := Enable, Reset := Reset, Causes := instCauses);
Fault := instFault.Fault;

ErrorEdge(CLK := Fault.Error);
IF ErrorEdge.Q AND NOT StepAtFaultCaptured THEN
    Outputs.StepAtFault := PrevState;
    StepAtFaultCaptured := TRUE;
ELSIF ResetEdge.Q AND NOT ErrorCausePresent AND NOT Inputs.KoboldImmersed
      AND NOT Inputs.MotionRequestActive AND NOT (Inputs.CurrentSpeedStep > 4) THEN
    Outputs.StepAtFault := E_DiveSearchState.WAIT_PRECONDITIONS;
END_IF;
{endregion}

{region "§2 Neutralisation et machine d'etat"}
IF NOT Enable OR NOT Inputs.PowerContactorEngaged THEN
    Ready := FALSE;
    Lifecycle.Busy := FALSE;
    Lifecycle.Done := FALSE;
    Outputs.DescendPermit := FALSE;
    Outputs.KoboldContactorCmd := FALSE;
    Outputs.BottomTouchConfirmed := FALSE;
    Outputs.StepState := E_DiveSearchState.WAIT_PRECONDITIONS;
    Outputs.OperatorActionId := 0;
    Outputs.OperatorAction := '';
    ImmersionConfirmed := FALSE;
    ImmersionTimerAcc := T#0ms;
    BottomTimerAcc := T#0ms;
    Outputs.MinStepDown := 0;
    PrevState := E_DiveSearchState.WAIT_PRECONDITIONS;
    RETURN;
END_IF;

Ready := Enable AND NOT Fault.Latched;
Outputs.DescendPermit := FALSE;
Outputs.KoboldContactorCmd := FALSE;
Lifecycle.Busy := FALSE;
Lifecycle.Done := FALSE;
Outputs.OperatorActionId := 0;
Outputs.OperatorAction := '';

DescentActive := Inputs.MotionRequestActive AND (Inputs.MotionDirection = -1)
              AND ((Inputs.Mode = E_Mode.MAINT_N1) OR (Inputs.Mode = E_Mode.MAINT_N2))
              AND NOT (Inputs.CurrentSpeedStep > 4)
              AND NOT SeqErrorFault;

IF Fault.Error OR Fault.Latched THEN
    Outputs.StepState := E_DiveSearchState.ERROR_HOLD;
    Outputs.KoboldContactorCmd := FALSE;
    Outputs.OperatorActionId := 16#0180;
    Outputs.OperatorAction := 'Verifier les conditions puis rearmer avant une nouvelle plongee.';
ELSE
    CASE Outputs.StepState OF
        E_DiveSearchState.WAIT_PRECONDITIONS:
            IF NOT Inputs.BypassPreconditions
               AND (NOT Inputs.BucketIsOpen OR NOT Inputs.PositionsValid OR Inputs.KoboldImmersed
                    OR (Inputs.M1Position_M < Inputs.DiveStartMin_M)
                    OR (Inputs.M2Position_M < Inputs.DiveStartMin_M)) THEN
                Outputs.OperatorActionId := 16#0100;
                Outputs.OperatorAction := 'Verifier benne ouverte, positions et Kobold au repos.';
            ELSE
                Outputs.StepState := E_DiveSearchState.READY_TO_DESCEND;
            END_IF;

        E_DiveSearchState.READY_TO_DESCEND:
            Ready := TRUE;
            Outputs.OperatorActionId := 16#0101;
            Outputs.OperatorAction := 'Demander une descente pour rechercher le fond.';
            IF Inputs.MotionRequestActive AND (Inputs.MotionDirection = -1) THEN
                ImmersionTimerAcc := T#0ms;
                Outputs.StepState := E_DiveSearchState.SEARCHING_IMMERSION;
            END_IF;

        E_DiveSearchState.SEARCHING_IMMERSION:
            Lifecycle.Busy := TRUE;
            Outputs.DescendPermit := DescentActive;
            Outputs.KoboldContactorCmd := DescentActive;
            Outputs.OperatorActionId := 16#0102;
            Outputs.OperatorAction := 'Maintenir la descente : recherche immersion Kobold.';
            IF Inputs.CurrentSpeedStep > 4 THEN
                IF NOT StepAtFaultCaptured THEN
                    Outputs.StepAtFault := Outputs.StepState;
                    StepAtFaultCaptured := TRUE;
                END_IF;
                Palier5ForbiddenFault := TRUE;
            END_IF;
            IF KoboldRiseEdge.Q THEN
                IF (Inputs.M1Position_M <= Inputs.ImmersionUpper_M)
                   AND (Inputs.M1Position_M >= Inputs.ImmersionLower_M)
                   AND (Inputs.M2Position_M <= Inputs.ImmersionUpper_M)
                   AND (Inputs.M2Position_M >= Inputs.ImmersionLower_M) THEN
                    ImmersionConfirmed := TRUE;
                    BottomTimerAcc := T#0ms;
                    Outputs.StepState := E_DiveSearchState.SEARCHING_BOTTOM;
                ELSE
                    IF NOT StepAtFaultCaptured THEN
                        Outputs.StepAtFault := Outputs.StepState;
                        StepAtFaultCaptured := TRUE;
                    END_IF;
                    SeqErrorFault := TRUE;
                END_IF;
            ELSIF (Inputs.M1Position_M < Inputs.ImmersionLower_M)
               OR (Inputs.M2Position_M < Inputs.ImmersionLower_M) THEN
                IF NOT StepAtFaultCaptured THEN
                    Outputs.StepAtFault := Outputs.StepState;
                    StepAtFaultCaptured := TRUE;
                END_IF;
                SeqErrorFault := TRUE;
            END_IF;

        E_DiveSearchState.SEARCHING_BOTTOM:
            Lifecycle.Busy := TRUE;
            Outputs.DescendPermit := DescentActive;
            Outputs.KoboldContactorCmd := DescentActive;
            Outputs.OperatorActionId := 16#0103;
            Outputs.OperatorAction := 'Maintenir la descente : immersion validee, recherche du fond.';
            IF Inputs.CurrentSpeedStep > 4 THEN
                IF NOT StepAtFaultCaptured THEN
                    Outputs.StepAtFault := Outputs.StepState;
                    StepAtFaultCaptured := TRUE;
                END_IF;
                Palier5ForbiddenFault := TRUE;
            END_IF;
            IF KoboldFallEdge.Q AND ImmersionConfirmed THEN
                Outputs.BottomTouchConfirmed := TRUE;
                ImmersionConfirmed := FALSE;
                Outputs.KoboldContactorCmd := FALSE;
                Outputs.StepState := E_DiveSearchState.BOTTOM_CONFIRMED;
            END_IF;

        E_DiveSearchState.BOTTOM_CONFIRMED:
            Lifecycle.Done := TRUE;
            Outputs.KoboldContactorCmd := FALSE;
            Outputs.OperatorActionId := 16#0104;
            Outputs.OperatorAction := 'Fond detecte : demander la fermeture ou extraction.';

        E_DiveSearchState.ERROR_HOLD:
            Outputs.KoboldContactorCmd := FALSE;
    END_CASE;
END_IF;

IF DescentActive AND ((Outputs.StepState = E_DiveSearchState.SEARCHING_IMMERSION)
                   OR (Outputs.StepState = E_DiveSearchState.SEARCHING_BOTTOM)) THEN
    Outputs.MinStepDown := LIMIT(0, Inputs.CfgDiveFloorStep, 5);
ELSE
    Outputs.MinStepDown := 0;
END_IF;

PrevState := Outputs.StepState;
{endregion}

END_FUNCTION_BLOCK

(* ---- FB_ExtractionAssist.st ---- *)
(* =======================================================================
   ⚙️ FB_ExtractionAssist — Fermeture benne et remontée assistée
   ───────────────────────────────────────────────────────────────
   🎯 Rôle : Séquence d'extraction (fermeture benne, remontée de contrôle, remontée nominale)
   🛡️ Sécurité : Aucune remontée assistée sans fond confirmé, contrôle palier 1
   📄 Doc métier : DOC/AF/AF_Partie-04_Mode_SemiAuto_Sequenceur_v2.3.md
   ======================================================================= *)
FUNCTION_BLOCK FB_ExtractionAssist
VAR_INPUT
    // === COMMANDES & AUTORISATIONS ===
    Enable                      : BOOL;     // --> [CMD] Activation generale du FB (TRUE=Autorise)
    Reset                       : BOOL;     // --> [CMD] Acquittement defaut (front)
    PowerContactorEngaged       : BOOL;     // --> [SAFE] Chaine de securite OK
    Mode                        : E_Mode;   // --> [CMD] Mode de fonctionnement arbitre
    MotionRequestActive         : BOOL;     // --> [CMD] Intention de mouvement active
    MotionDirection             : INT;      // --> [CMD] Sens de mouvement (+1 = montee)
    BottomPositionConfirmed     : BOOL;     // --> [SAFE] Attestation fond confirme (Kobold ou op)

    // === CAPTEURS & ETATS MATERIELS ===
    BucketIsClosed              : BOOL;     // --> [HW] Benne fermee confirmee
    BucketBusy                  : BOOL;     // --> [HW] Mouvement benne en cours
    BucketError                 : BOOL;     // --> [SAFE] Defaut sur sous-systeme benne
    WinchSyncError              : BOOL;     // --> [SAFE] Defaut de desynchronisme treuils M1/M2
    M1Position_M                : REAL;     // --> [HW] Position codeur treuil M1 (m)
    M2Position_M                : REAL;     // --> [HW] Position codeur treuil M2 (m)
    M1MeasuredSpeedValid        : BOOL;     // --> [HW] Validite mesure vitesse M1
    M2MeasuredSpeedValid        : BOOL;     // --> [HW] Validite mesure vitesse M2
    PositionsValid              : BOOL;     // --> [HW] Validite des mesures de position

    // === CONFIGURATION & REGLAGES ===
    ControlAscentDistance_M     : REAL;     // --> [CFG] Distance palier 1 de controle remontee (m)
    CfgBucketCloseTimeout       : TIME := T#75s;// --> [CFG] Backstop fermeture benne (doit rester > BucketMoveTimeout)
    BucketMoveTimeout           : TIME := T#60s;// --> [CFG] Reference watchdog mouvement FB_Bucket (verrouillage ordre backstop)
    CycleTime                   : TIME := T#10ms;// --> [CFG] Base de temps d'integration (periode MainTask)
END_VAR
VAR_OUTPUT
    // === ETATS IEC & DEFECTUOSITES ===
    Ready                       : BOOL;     // <-- [STAT] FB pret a fonctionner
    // 🧩 Statut transverse (forme cible ST_Fault + ST_Lifecycle)
    Fault                       : ST_Fault;
    Lifecycle                   : ST_Lifecycle;
    ExtractionState             : E_ExtractionAssistState; // <-- [STAT] Phase interne extraction
    StepAtFault                 : E_ExtractionAssistState; // <-- [DIAG] Phase active memorisee lors du defaut

    // === ORDRES & AUTORISATIONS ===
    BucketCloseRequest          : BOOL;     // <-- [ACT] Demande de fermeture benne
    AscentPermit                : BOOL;     // <-- [ACT] Autorisation de remontee assistee
    ExtractionControlActive     : BOOL;     // <-- [ACT] Plafond palier 1 pendant la montee controlee
    BottomConfirmationConsumed  : BOOL;     // <-- [STAT] Signal confirmation fond consomme

    // === DIAGNOSTIC IHM ===
    OperatorActionId            : WORD;     // <-- [DIAG] ID action operateur requise
    OperatorAction              : STRING(120); // <-- [DIAG] Message explicatif operateur
END_VAR
VAR
    // === DETECTEURS DE FRONTS ===
    ResetEdge                   : R_TRIG;   // . [LOC] Detecteur front montant Reset
    ErrorEdge                   : R_TRIG;   // . [LOC] Detecteur front montant apparition defaut

    // === MEMORISATIONS & POSITIONS INTERNES ===
    ControlStartM1Position_M    : REAL;     // . [LOC] Position M1 au debut du palier de controle (m)
    ControlStartM2Position_M    : REAL;     // . [LOC] Position M2 au debut du palier de controle (m)
    PrevState                   : E_ExtractionAssistState; // . [LOC] Phase au scan precedent (survit au gate)

    // === CALCUL DYNAMIQUE RUNTIME DU TIMEOUT DECOLLAGE ===
    CalculatedControlAscentTimeout : TIME;  // . [LOC] Plafond anti-blocage decollage calcule au runtime

    // === ACCUMULATEURS DE TEMPS ANTI-POMPAGE ===
    BucketCloseTimerAcc         : TIME := T#0ms;// . [LOC] Temps cumule fermeture benne sous montee demandee
    ControlAscentTimerAcc       : TIME := T#0ms;// . [LOC] Temps cumule decollage controle sous montee demandee

    // === VARIABLES LOCALES INTERNES ===
    ErrorCausePresent           : BOOL;     // . [LOC] Presence d'une cause de defaut parametrage
    BucketErrorFault            : BOOL;     // . [LOC] Latch erreur benne
    SyncOrSpeedErrorFault       : BOOL;     // . [LOC] Latch erreur synchro/vitesse
    TimeoutBucketCloseFault     : BOOL;     // . [LOC] Latch backstop fermeture benne
    TimeoutControlAscentFault   : BOOL;     // . [LOC] Latch timeout decollage controle
    StepAtFaultCaptured         : BOOL;     // . [LOC] StepAtFault deja fige pour l'episode de defaut courant
    AssistPermit                : BOOL;     // . [LOC] Ascending assistee reellement demandee (sens + mode)
    AscentControlSafe           : BOOL;     // . [LOC] Entrees [SAFE] saines pour le decollage controle
    AscentNominalSafe           : BOOL;     // . [LOC] Entrees [SAFE] saines pour la remontee nominale
    CausesPhysiquesEffacees     : BOOL;     // . [LOC] Toutes les entrees defaut treuil/benne revenues a l'etat sain

    // === SOCLE DEFAUT ===
    instFault                   : FB_FaultCore;                  // * [INST] Socle défaut transverse
    instCauses                  : ARRAY[0..15] OF ST_FaultCause; // . [LOC] Table des causes nommées
END_VAR
VAR CONSTANT
    // === CONSTANTES DERIVATION TIMEOUT ANTI-BLOCAGE ===
    CST_MinSpeed_Mps            : REAL := 0.15;   // Vitesse Palier 1 mini sous charge/mou (m/s)
    CST_ControlAscentMargin     : REAL := 2.0;    // Facteur de marge sur la course de decollage
    CST_TimeoutMinDistance_M    : REAL := 0.1;    // Plancher de distance pour le calcul (evite timeout degenere)
    CST_TimeoutMaxDistance_M    : REAL := 20.0;   // Plafond de distance : borne le calcul avant REAL_TO_UDINT (anti-overflow)
    CST_BackstopMax             : TIME := T#600s; // Plafond du backstop fermeture benne : au-dela, risque d'overflow de l'accumulateur
    CST_SecToMs                 : REAL := 1000.0; // Conversion secondes -> millisecondes
END_VAR

// === IMPLEMENTATION ===

{region "§1 Causes & Socle Défaut (évalué en continu)"}
// 🔑 1. FRONTS
ResetEdge(CLK := Reset);
// Parametrage invalide : distance nulle, backstop nul, base de temps nulle, ou backstop
// qui fauterait AVANT le watchdog benne (masquerait BucketError - ordre des watchdogs).
ErrorCausePresent := (ControlAscentDistance_M <= 0.0)
                  OR (CfgBucketCloseTimeout <= T#0ms)
                  OR (CycleTime <= T#0ms)
                  OR (CfgBucketCloseTimeout <= BucketMoveTimeout)
                  OR (CfgBucketCloseTimeout > CST_BackstopMax);  // borne haute : evite l'overflow de BucketCloseTimerAcc (F3)

// ⏱️ Plafond anti-blocage decollage calcule au runtime : course de controle bornee [plancher..plafond]
// avant conversion REAL->UDINT->TIME (anti-overflow sur valeur IHM aberrante, CQS §6).
CalculatedControlAscentTimeout := UDINT_TO_TIME(REAL_TO_UDINT(
    LIMIT(CST_TimeoutMinDistance_M, ControlAscentDistance_M, CST_TimeoutMaxDistance_M)
    / CST_MinSpeed_Mps * CST_ControlAscentMargin * CST_SecToMs));

// ⏱️ Integrateurs de temps de montee effective (anti-pompage homme-mort)
IF (ExtractionState = E_ExtractionAssistState.CLOSING_BUCKET) AND MotionRequestActive AND (MotionDirection = 1) THEN
    BucketCloseTimerAcc := BucketCloseTimerAcc + CycleTime;
    IF BucketCloseTimerAcc >= CfgBucketCloseTimeout THEN
        TimeoutBucketCloseFault := TRUE;
    END_IF;
END_IF;

IF (ExtractionState = E_ExtractionAssistState.CONTROL_ASCENT) AND MotionRequestActive AND (MotionDirection = 1) THEN
    ControlAscentTimerAcc := ControlAscentTimerAcc + CycleTime;
    IF ControlAscentTimerAcc >= CalculatedControlAscentTimeout THEN
        TimeoutControlAscentFault := TRUE;
    END_IF;
END_IF;

// Etat physique des causes treuil/benne : conditionne l'acquittement des latches a cause persistante (F2).
CausesPhysiquesEffacees := NOT BucketError AND NOT WinchSyncError
                        AND PositionsValid AND M1MeasuredSpeedValid AND M2MeasuredSpeedValid;
IF ResetEdge.Q AND NOT ErrorCausePresent AND NOT MotionRequestActive THEN
    // Latches sans cause physique persistante (timeouts, backstop) : acquittables sur simple front Reset.
    TimeoutBucketCloseFault   := FALSE;
    TimeoutControlAscentFault := FALSE;
    BucketCloseTimerAcc       := T#0ms;
    ControlAscentTimerAcc     := T#0ms;
    StepAtFaultCaptured       := FALSE;
    ExtractionState := E_ExtractionAssistState.WAIT_BOTTOM_CONFIRMATION;
    // Latches de cause physique : acquittables SEULEMENT si l'entree de defaut est revenue saine (F2).
    IF CausesPhysiquesEffacees THEN
        BucketErrorFault      := FALSE;
        SyncOrSpeedErrorFault := FALSE;
    END_IF;
END_IF;

instCauses[1].Active   := BucketErrorFault;
instCauses[1].Latching := TRUE;
instCauses[1].Texte    := 'Defaut sous-systeme benne pendant fermeture';

instCauses[2].Active   := SyncOrSpeedErrorFault;
instCauses[2].Latching := TRUE;
instCauses[2].Texte    := 'Defaut synchro ou capteurs treuils pendant remontee';

instCauses[3].Active   := ErrorCausePresent;
instCauses[3].Latching := TRUE;
instCauses[3].Texte    := 'Parametrage distance de controle ou backstop invalide';

instCauses[4].Active   := TimeoutBucketCloseFault;
instCauses[4].Latching := TRUE;
instCauses[4].Texte    := 'Depassement backstop fermeture benne';

instCauses[5].Active   := TimeoutControlAscentFault;
instCauses[5].Latching := TRUE;
instCauses[5].Texte    := 'Depassement tempo decollage controle';

// Appel du socle de défaut
instFault(Enable := Enable, Reset := Reset, Causes := instCauses);
Fault := instFault.Fault;

// 📸 Capture ordonnee de StepAtFault (D2). Les defauts leves dans le CASE se figent au site du
// latch (voir §3) ; ce bloc ne couvre que les defauts detectes en §1 (backstop, timeout, parametrage),
// ou ExtractionState/PrevState sont encore l'etape reelle. StepAtFaultCaptured evite l'ecrasement.
ErrorEdge(CLK := Fault.Error);
IF ErrorEdge.Q AND NOT StepAtFaultCaptured THEN
    StepAtFault := PrevState;
    StepAtFaultCaptured := TRUE;
ELSIF ResetEdge.Q AND NOT ErrorCausePresent AND NOT MotionRequestActive THEN
    StepAtFault := E_ExtractionAssistState.WAIT_BOTTOM_CONFIRMATION;
END_IF;
{endregion}

{region "§2 Gate neutralisation"}
// 🛑 2. GATE
IF NOT Enable OR NOT PowerContactorEngaged THEN
    Ready := FALSE;
    Lifecycle.Busy := FALSE;
    Lifecycle.Done := FALSE;
    BucketCloseRequest := FALSE;
    AscentPermit := FALSE;
    ExtractionControlActive := FALSE;
    BottomConfirmationConsumed := FALSE;
    ExtractionState := E_ExtractionAssistState.WAIT_BOTTOM_CONFIRMATION;
    // StepAtFault / StepAtFaultCaptured NON reinitialises ici : l'etape figee au defaut reste
    // lisible pour l'IHM/diagnostic apres un cycle Enable OFF->ON ; seul un front Reset l'efface.
    PrevState := E_ExtractionAssistState.WAIT_BOTTOM_CONFIRMATION;
    BucketCloseTimerAcc := T#0ms;
    ControlAscentTimerAcc := T#0ms;
    OperatorActionId := 0;
    OperatorAction := '';
    RETURN;
END_IF;

Ready := Enable AND NOT Fault.Latched;
{endregion}

{region "§3 Machine etat fermeture remontee"}
BucketCloseRequest := FALSE;
AscentPermit := FALSE;
ExtractionControlActive := FALSE;
BottomConfirmationConsumed := FALSE;
Lifecycle.Busy := FALSE;
Lifecycle.Done := FALSE;

// Ascending assistee reellement demandee : sens ascending + mode maintenance (H5, double garde vs Enable PRG_03).
AssistPermit := MotionRequestActive AND (MotionDirection = 1)
            AND (Mode = E_Mode.MAINT_N1 OR Mode = E_Mode.MAINT_N2);
// Entrees [SAFE] saines : coupure meme-scan des permis si defaut treuil/synchro (H2), avant meme le latch.
AscentControlSafe := NOT WinchSyncError AND PositionsValid AND M1MeasuredSpeedValid AND M2MeasuredSpeedValid;
AscentNominalSafe := NOT WinchSyncError AND PositionsValid;

// Garde-fou non-redemarrage auto : un defaut latche non acquitte verrouille la machine
// d'etat en ERROR_HOLD, meme si la vue live Fault.Error retombe (cause disparue).
IF Fault.Error OR Fault.Latched THEN
    ExtractionState := E_ExtractionAssistState.ERROR_HOLD;
    OperatorActionId := 16#0280;
    OperatorAction := 'Vérifier la benne et les treuils puis réarmer avant de reprendre.';
ELSE
    CASE ExtractionState OF
        E_ExtractionAssistState.WAIT_BOTTOM_CONFIRMATION:
            IF BottomPositionConfirmed THEN
                ExtractionState := E_ExtractionAssistState.READY_TO_CLOSE;
            ELSE
                OperatorActionId := 16#0200;
                OperatorAction := 'Confirmer que la benne est posée au fond avant extraction.';
            END_IF;

        E_ExtractionAssistState.READY_TO_CLOSE:
            Ready := TRUE;
            OperatorActionId := 16#0201;
            OperatorAction := 'Demander la montée pour fermer la benne.';
            IF MotionRequestActive AND (MotionDirection = 1) THEN
                BottomConfirmationConsumed := TRUE;
                BucketCloseTimerAcc := T#0ms;   // ⏱️ RAZ a l'entree exacte de CLOSING_BUCKET
                ExtractionState := E_ExtractionAssistState.CLOSING_BUCKET;
            END_IF;

        E_ExtractionAssistState.CLOSING_BUCKET:
            Lifecycle.Busy := TRUE;
            BucketCloseRequest := AssistPermit AND NOT BucketError; // coupure meme-scan sur defaut benne (H2)
            // Autorisation de montee pendant la fermeture : la benne se ferme en montant.
            // Consommee par l'arbitrage (PRG_04) comme permis de montee assistee (H2).
            AscentPermit := AssistPermit AND AscentControlSafe;
            OperatorActionId := 16#0202;
            OperatorAction := 'Maintenir la montée : fermeture de la benne en cours.';
            IF BucketError THEN
                IF NOT StepAtFaultCaptured THEN
                    StepAtFault := ExtractionState;
                    StepAtFaultCaptured := TRUE;
                END_IF;
                BucketErrorFault := TRUE;
            ELSIF BucketIsClosed AND NOT BucketBusy THEN
                ControlStartM1Position_M := M1Position_M;
                ControlStartM2Position_M := M2Position_M;
                ControlAscentTimerAcc := T#0ms;   // ⏱️ RAZ a l'entree exacte de CONTROL_ASCENT
                ExtractionState := E_ExtractionAssistState.CONTROL_ASCENT;
            END_IF;

        E_ExtractionAssistState.CONTROL_ASCENT:
            Lifecycle.Busy := TRUE;
            AscentPermit := AssistPermit AND AscentControlSafe; // coupure meme-scan sur defaut synchro/capteurs (H2)
            ExtractionControlActive := AscentPermit;            // plafond palier 1 suit le permis de montee
            OperatorActionId := 16#0203;
            OperatorAction := 'Maintenir la montée : contrôle charge au palier minimal.';
            IF NOT AscentControlSafe THEN
                IF NOT StepAtFaultCaptured THEN
                    StepAtFault := ExtractionState;
                    StepAtFaultCaptured := TRUE;
                END_IF;
                SyncOrSpeedErrorFault := TRUE;
            ELSIF (M1Position_M >= (ControlStartM1Position_M + ControlAscentDistance_M))
               AND (M2Position_M >= (ControlStartM2Position_M + ControlAscentDistance_M)) THEN
                ExtractionState := E_ExtractionAssistState.NOMINAL_ASCENT;
            END_IF;

        E_ExtractionAssistState.NOMINAL_ASCENT:
            Lifecycle.Busy := TRUE;
            AscentPermit := AssistPermit AND AscentNominalSafe; // coupure meme-scan sur defaut synchro/position (H2)
            OperatorActionId := 16#0204;
            OperatorAction := 'Maintenir la montée : extraction en cours.';
            IF NOT AscentNominalSafe THEN
                IF NOT StepAtFaultCaptured THEN
                    StepAtFault := ExtractionState;
                    StepAtFaultCaptured := TRUE;
                END_IF;
                SyncOrSpeedErrorFault := TRUE;
            END_IF;

        E_ExtractionAssistState.ERROR_HOLD:
            ;
    END_CASE;
END_IF;

// 💾 Memorisation de la phase precedente en toute fin de scan (capture StepAtFault fiable)
PrevState := ExtractionState;
{endregion}

END_FUNCTION_BLOCK

(* ---- FB_MachineHomingCycle.st ---- *)
(* =======================================================================
   🎯 FB_MachineHomingCycle — Guide de referencement machine M1/M2/benne
   ───────────────────────────────────────────────────────────────
   🎯 Role : Qualifier le datum machine (2 codeurs cales + etat benne
             confirme) et guider le homing conjoint M1/M2 + le commit
             atomique de l'etat benne. N'emet AUCUN ordre de mouvement.
   🔒 Securite : SEMI_AUTO interdit tant que MachineHomed=FALSE. Perte de
                 datum en mouvement -> SafeStop ; reprise sur Reset conscient
                 uniquement (aucun redemarrage automatique).
   🔌 Interface : contrat standard (Enable/Reset, Ready/Fault/Lifecycle).
                  Producteur UNIQUE de la qualification machine — ne relit
                  jamais un ActiveOffsetValid aval (C).
   📄 Doc metier : DOC/AF/AF_Partie-09_Fonction_Encoder_v2.4.md (F09.08)
                   + DOC/AF/AF_Partie-05_Modes_Maintenance_v2.1.md
   🧩 Dependances : FB_FaultCore, FB_Encoder (M1/M2), FB_Bucket, FB_Modes
   ======================================================================= *)
FUNCTION_BLOCK PUBLIC FB_MachineHomingCycle
VAR_INPUT
    // === CONTRAT STANDARD (Enable + Reset) ===
    Enable                      : BOOL;                                      // --> [CMD] Autorisation generale (FALSE => sorties sures, retour IDLE)
    Reset                       : BOOL;                                      // --> [CMD] Acquittement defaut (front, jamais conditionne)

    // === MODE ARBITRE ===
    Mode                        : E_Mode;                                    // --> [CMD] Mode machine (confirmation benne : MAINT_N2 seul)

    // === PERMIS SECURITE ===
    TopPositionActive           : BOOL;                                      // --> [SAFE] Capteur haut commun au contact
    WinchesMechanicallyStopped  : BOOL;                                      // --> [SAFE] M1 ET M2 arret mecanique confirme

    // === ACQUISITION HOMING (M1 / M2) ===
    M1Status                    : ST_fbMachineHomingCycle_AxisHomingStatus;  // --> [HW] Statut homing axe M1 (Retenue)
    M2Status                    : ST_fbMachineHomingCycle_AxisHomingStatus;  // --> [HW] Statut homing axe M2 (Benne)

    // === ETAT BENNE ===
    BucketOffsetValid           : BOOL;                                      // --> [HW] Offset benne actif valide (FB_Bucket) — bootstrap datum seulement

    // === COMMANDES OPERATEUR (IHM) ===
    ConfirmOpenPosition         : BOOL;                                      // --> [CMD] Confirmation visuelle "benne ouverte" (niveau, front interne)
    ConfirmClosePosition        : BOOL;                                      // --> [CMD] Confirmation visuelle "benne fermee" (niveau, front interne)

    // === REGLAGES & CONFIGURATION ===
    Cfg                         : ST_fbMachineHomingCycle_Cfg;              // --> [CFG] Reglages geometriques referencement (cible M1 + ecarts benne)
END_VAR
VAR_OUTPUT
    // === CONTRAT STANDARD (Ready + Fault) ===
    Ready                       : BOOL;                                      // <-- [STAT] FB actif (Enable ET NOT Fault.Latched)
    Fault                       : ST_Fault;                                  // <-- [SAFE] Socle defaut (rempli par FB_FaultCore)
    Lifecycle                   : ST_Lifecycle;                              // <-- [STAT] Cycle transaction (Busy = homing conjoint en cours)

    // === QUALIFICATION MACHINE ===
    MachineHomed                : BOOL;                                      // <-- [SAFE] Datum machine valide (gate SEMI_AUTO)
    MachineHomingStep           : E_MachineHomingStep := E_MachineHomingStep.IDLE;   // <-- [STAT] Etape du guide
    MachineHomingStepAtError    : E_MachineHomingStep := E_MachineHomingStep.IDLE;   // <-- [DIAG] Etape figee a l'apparition du defaut (R9)
    MachineHomingInstruction    : STRING(120);                              // <-- [DIAG] Consigne operateur en clair (ASCII)
    MachineHomingActive         : BOOL;                                      // <-- [STAT] Transaction en cours (= Lifecycle.Busy)
    MachineHomingLossSafeStop   : BOOL;                                      // <-- [SAFE] Demande d'arret controle suite perte de datum en mouvement
    MachineHomingFailed         : BOOL;                                      // <-- [STAT] Derniere transaction abandonnee

    // === DEMANDES HOMING (M1 / M2) ===
    M1Demand                    : ST_fbMachineHomingCycle_HomingDemand;      // <-- [ACT] Demande de homing conjoint axe M1
    M2Demand                    : ST_fbMachineHomingCycle_HomingDemand;      // <-- [ACT] Demande de homing conjoint axe M2 (cible dynamique)

    // === COMMIT BENNE ===
    BucketCommit                : ST_fbMachineHomingCycle_BucketCommit;      // <-- [ACT] Publication atomique de l'etat benne (vers FB_Bucket)
END_VAR
VAR
    // === SOUS-INSTANCES FB ===
    instFault                   : FB_FaultCore;                             // * [INST] Socle defaut transverse
    ResetEdge                   : R_TRIG;                                   // * [INST] Front montant Reset
    ConfirmOpenEdge             : R_TRIG;                                   // * [INST] Front montant ConfirmOpenPosition
    ConfirmCloseEdge            : R_TRIG;                                   // * [INST] Front montant ConfirmClosePosition
    LatchedEdge                 : R_TRIG;                                   // * [INST] Front montant Fault.Latched (capture R9)

    // === TABLE DES CAUSES DE DEFAUT ===
    instCauses                  : ARRAY[0..15] OF ST_FaultCause;            // . [LOC] Causes en clair pour FB_FaultCore

    // === ETATS INTERNES TRANSACTION ===
    PendingOpen                 : BOOL;                                     // . [LOC] Confirmation "ouverte" en attente de commit
    PendingClose                : BOOL;                                     // . [LOC] Confirmation "fermee" en attente de commit
    HomingStarted               : BOOL;                                     // . [LOC] Transaction homing conjoint armee
    HomingBusyObserved          : BOOL;                                     // . [LOC] Au moins un Busy observe depuis le debut de la transaction
    CommitPublished             : BOOL;                                     // . [LOC] Commit benne deja publie sur ce datum
    MachineWasHomed             : BOOL;                                     // . [LOC] Memorise un datum valide (detection de perte)
    HomingLossLatched           : BOOL;                                     // . [LOC] Perte de datum en mouvement latchee jusqu'a l'arret
    ReHomingAckRequired         : BOOL;                                     // . [LOC] C-1 : bloque MachineHomed jusqu'a un Reset conscient

    // === CONDITIONS INTERMEDIAIRES NOMMEES (std 2quater : <= 3 termes) ===
    DoubleConfirmRequested      : BOOL;                                     // . [LOC] Les deux fronts confirmation au meme scan (C-2)
    SingleConfirm               : BOOL;                                     // . [LOC] Exactement un front confirmation
    ConfirmWhileHoming          : BOOL;                                     // . [LOC] Confirmation pendant un homing d'axe en cours (C-4.3)
    WindowSafe                  : BOOL;                                     // . [LOC] Fenetre mecanique sure (N2 + capteur haut + arret)
    AxisHomed                   : BOOL;                                     // . [LOC] M1 ET M2 references et fiables
    CommitOrOffsetValid         : BOOL;                                     // . [LOC] Datum benne connu (commit publie OU offset valide)
    TransactionAbort            : BOOL;                                     // . [LOC] Condition d'abandon fail-safe de la transaction
    MachineHomedRaw             : BOOL;                                     // . [LOC] Qualification hors Fault (detection de perte, evite la circularite)
END_VAR
VAR CONSTANT
    // === INDICES DE CAUSES (instCauses[]) ===
    CST_CAUSE_HOMING_LOST_IN_MOTION : INT := 0;                             // Perte d'un datum valide pendant un mouvement (Latching)
    CST_CAUSE_TX_ABORT_TOP_LOST     : INT := 1;                             // Capteur haut perdu pendant la transaction (Latching)
    CST_CAUSE_TX_ABORT_MOTION       : INT := 2;                             // Mouvement detecte pendant la transaction (Latching)
    CST_CAUSE_HOMING_ERROR_M1       : INT := 3;                             // FB_Encoder M1 signale une erreur de homing (Latching)
    CST_CAUSE_HOMING_ERROR_M2       : INT := 4;                             // FB_Encoder M2 signale une erreur de homing (Latching)
    CST_CAUSE_DOUBLE_CONFIRM        : INT := 5;                             // ConfirmOpen ET ConfirmClose au meme scan (Latching) — C-2
    CST_CAUSE_CONFIRM_WHILE_HOMING  : INT := 6;                             // Confirmation pendant un homing d'axe en cours (Latching) — C-4.3
END_VAR

// === 🔑 §1 FRONTS, CIBLE DYNAMIQUE, CAUSES ET SOCLE DEFAUT ===
{region "§1 Fronts & causes"}

// Sorties impulsionnelles remises a FALSE en tete de scan (1 scan actif au commit / a la demande).
M1Demand.HomeReq := FALSE;
M2Demand.HomeReq := FALSE;
BucketCommit.CommitOpen := FALSE;
BucketCommit.CommitClose := FALSE;

// Cible dynamique M2 : recalculee chaque scan (jamais une position M1 live).
M2Demand.UseDynamicTarget := PendingOpen OR PendingClose OR HomingStarted;
IF PendingClose THEN
    M2Demand.DynamicTarget_M := Cfg.CfgTopHomingTarget_M + Cfg.CfgOffsetClose_M;
ELSE
    M2Demand.DynamicTarget_M := Cfg.CfgTopHomingTarget_M + Cfg.CfgOffsetOpen_M;
END_IF;
M1Demand.UseDynamicTarget := FALSE;

// Detection de fronts.
ResetEdge(CLK := Reset);
ConfirmOpenEdge(CLK := ConfirmOpenPosition);
ConfirmCloseEdge(CLK := ConfirmClosePosition);
LatchedEdge(CLK := Fault.Latched);

// Purge sur front Reset (inclut C-1 : ReHomingAckRequired).
IF ResetEdge.Q THEN
    PendingOpen         := FALSE;
    PendingClose        := FALSE;
    HomingStarted       := FALSE;
    HomingBusyObserved  := FALSE;
    CommitPublished     := FALSE;
    MachineHomingFailed := FALSE;
    MachineWasHomed     := FALSE;
    HomingLossLatched   := FALSE;
    ReHomingAckRequired := FALSE;
END_IF;

// Conditions intermediaires nommees (std 2quater).
DoubleConfirmRequested := ConfirmOpenEdge.Q AND ConfirmCloseEdge.Q;
SingleConfirm          := ConfirmOpenEdge.Q XOR ConfirmCloseEdge.Q;
ConfirmWhileHoming     := SingleConfirm AND (M1Status.HomingBusy OR M2Status.HomingBusy);
WindowSafe             := (Mode = E_Mode.MAINT_N2) AND TopPositionActive AND WinchesMechanicallyStopped;
AxisHomed              := M1Status.HomedAndReliable AND M2Status.HomedAndReliable;
CommitOrOffsetValid    := CommitPublished OR BucketOffsetValid;

// Qualification "brute" (sans Fault) : sert a la detection de perte sans creer de circularite
// avec le socle defaut appele plus bas.
MachineHomedRaw := AxisHomed AND CommitOrOffsetValid
                   AND NOT MachineHomingFailed AND NOT ReHomingAckRequired;

// Perte d'un datum auparavant valide EN MOUVEMENT : latch jusqu'a l'arret mecanique.
IF MachineHomedRaw THEN
    MachineWasHomed := TRUE;
END_IF;
IF MachineWasHomed AND NOT MachineHomedRaw AND NOT WinchesMechanicallyStopped THEN
    HomingLossLatched := TRUE;
END_IF;
IF NOT MachineHomedRaw AND WinchesMechanicallyStopped THEN
    MachineWasHomed := FALSE;
END_IF;
IF HomingLossLatched AND WinchesMechanicallyStopped THEN
    HomingLossLatched := FALSE;
END_IF;

(* C : pas de redemarrage automatique. Une perte de datum en mouvement exige un
   acquittement conscient (front Reset) avant que MachineHomed puisse revenir. *)
IF HomingLossLatched AND NOT ReHomingAckRequired THEN
    ReHomingAckRequired := TRUE;
END_IF;

// Table des causes (toutes Latching : acquittables au front Reset).
instCauses[CST_CAUSE_HOMING_LOST_IN_MOTION].Active   := HomingLossLatched OR ReHomingAckRequired;
instCauses[CST_CAUSE_HOMING_LOST_IN_MOTION].Latching := TRUE;
instCauses[CST_CAUSE_HOMING_LOST_IN_MOTION].Texte    := 'Perte de datum machine en mouvement : re-referencer';

instCauses[CST_CAUSE_TX_ABORT_TOP_LOST].Active   := HomingStarted AND NOT TopPositionActive;
instCauses[CST_CAUSE_TX_ABORT_TOP_LOST].Latching := TRUE;
instCauses[CST_CAUSE_TX_ABORT_TOP_LOST].Texte    := 'Capteur haut perdu pendant le referencement conjoint';

instCauses[CST_CAUSE_TX_ABORT_MOTION].Active   := HomingStarted AND NOT WinchesMechanicallyStopped;
instCauses[CST_CAUSE_TX_ABORT_MOTION].Latching := TRUE;
instCauses[CST_CAUSE_TX_ABORT_MOTION].Texte    := 'Mouvement detecte pendant le referencement conjoint';

instCauses[CST_CAUSE_HOMING_ERROR_M1].Active   := HomingStarted AND M1Status.HomingError;
instCauses[CST_CAUSE_HOMING_ERROR_M1].Latching := TRUE;
instCauses[CST_CAUSE_HOMING_ERROR_M1].Texte    := 'Erreur de homing codeur M1 pendant le referencement conjoint';

instCauses[CST_CAUSE_HOMING_ERROR_M2].Active   := HomingStarted AND M2Status.HomingError;
instCauses[CST_CAUSE_HOMING_ERROR_M2].Latching := TRUE;
instCauses[CST_CAUSE_HOMING_ERROR_M2].Texte    := 'Erreur de homing codeur M2 pendant le referencement conjoint';

(* C : confirmation Ouverte ET Fermee au meme scan = rejet total, cause a acquitter. *)
instCauses[CST_CAUSE_DOUBLE_CONFIRM].Active   := DoubleConfirmRequested;
instCauses[CST_CAUSE_DOUBLE_CONFIRM].Latching := TRUE;
instCauses[CST_CAUSE_DOUBLE_CONFIRM].Texte    := 'Confirmation benne Ouverte et Fermee simultanee : refusee';

(* C : confirmation recue pendant un homing d'axe deja en cours = ignoree. *)
instCauses[CST_CAUSE_CONFIRM_WHILE_HOMING].Active   := ConfirmWhileHoming;
instCauses[CST_CAUSE_CONFIRM_WHILE_HOMING].Latching := TRUE;
instCauses[CST_CAUSE_CONFIRM_WHILE_HOMING].Texte    := 'Confirmation benne pendant un homing codeur en cours : ignoree';

// Socle defaut : appele AVANT la gate NOT Enable (Reset jamais conditionne, std 9).
instFault(Enable := Enable, Reset := Reset, Causes := instCauses);
Fault := instFault.Fault;
{endregion}

// === 🔑 §2 DEMANDE SAFESTOP SUR PERTE DE DATUM ===
{region "§2 Perte datum"}
// Demande d'arret controle tant que la perte n'est pas mecaniquement resolue.
// La qualification de sortie MachineHomed est calculee en §6, APRES le deroule de
// transaction (commit ou abandon du meme scan pris en compte) — calcul unique.
MachineHomingLossSafeStop := HomingLossLatched;
{endregion}

// === 🔑 §3 GATE D'INITIALISATION (NOT Enable) ===
{region "§3 Gate init NOT Enable"}
IF NOT Enable THEN
    MachineHomingStep         := E_MachineHomingStep.IDLE;
    MachineHomingInstruction  := 'Referencement indisponible';
    MachineHomed              := FALSE;
    MachineHomingActive       := FALSE;
    M1Demand.HomeReq          := FALSE;
    M2Demand.HomeReq          := FALSE;
    M1Demand.UseDynamicTarget := FALSE;
    M2Demand.UseDynamicTarget := FALSE;
    BucketCommit.CommitOpen   := FALSE;
    BucketCommit.CommitClose  := FALSE;
    Lifecycle.Busy            := FALSE;
    Lifecycle.Done            := FALSE;
    Ready                     := FALSE;
    RETURN;
END_IF;
{endregion}

// === 🔑 §4 OUVERTURE DE LA TRANSACTION DE REFERENCEMENT CONJOINT ===
{region "§4 Ouverture transaction"}
(* C : jamais "au vol" par-dessus un homing d'axe deja en cours.
   Demande acceptee uniquement dans la fenetre mecanique sure, front unique, hors double. *)
IF SingleConfirm AND NOT HomingStarted AND NOT DoubleConfirmRequested AND NOT ConfirmWhileHoming
   AND WindowSafe
   AND NOT M1Status.HomingBusy AND NOT M2Status.HomingBusy THEN
    PendingOpen        := ConfirmOpenEdge.Q;
    PendingClose       := ConfirmCloseEdge.Q;
    HomingStarted      := TRUE;
    HomingBusyObserved := FALSE;
    CommitPublished    := FALSE;
    MachineHomingFailed := FALSE;
    M1Demand.HomeReq          := TRUE;
    M2Demand.HomeReq          := TRUE;
    M2Demand.UseDynamicTarget := TRUE;
    IF PendingClose THEN
        M2Demand.DynamicTarget_M := Cfg.CfgTopHomingTarget_M + Cfg.CfgOffsetClose_M;
    ELSE
        M2Demand.DynamicTarget_M := Cfg.CfgTopHomingTarget_M + Cfg.CfgOffsetOpen_M;
    END_IF;
END_IF;
{endregion}

// === 🔑 §5 DEROULE DE LA TRANSACTION & COMMIT ATOMIQUE ===
{region "§5 Deroule transaction & commit atomique"}
IF HomingStarted THEN
    M2Demand.UseDynamicTarget := TRUE;
    IF PendingClose THEN
        M2Demand.DynamicTarget_M := Cfg.CfgTopHomingTarget_M + Cfg.CfgOffsetClose_M;
    ELSE
        M2Demand.DynamicTarget_M := Cfg.CfgTopHomingTarget_M + Cfg.CfgOffsetOpen_M;
    END_IF;

    TransactionAbort := (NOT TopPositionActive) OR (NOT WinchesMechanicallyStopped)
                        OR M1Status.HomingError OR M2Status.HomingError;

    IF TransactionAbort THEN
        MachineHomingFailed := TRUE;
        HomingStarted       := FALSE;
        PendingOpen         := FALSE;
        PendingClose        := FALSE;
    ELSIF M1Status.HomingBusy OR M2Status.HomingBusy THEN
        HomingBusyObserved := TRUE;
    ELSIF HomingBusyObserved AND M1Status.HomedAndReliable AND M2Status.HomedAndReliable
          AND M1Status.HomingDone AND M2Status.HomingDone THEN
        (* Publication atomique : les deux etats benne ecrits par FB_Bucket dans le meme
           scan, uniquement apres les deux succes observes. *)
        BucketCommit.CommitOpen  := PendingOpen;
        BucketCommit.CommitClose := PendingClose;
        CommitPublished := TRUE;
        HomingStarted   := FALSE;
        PendingOpen     := FALSE;
        PendingClose    := FALSE;
    END_IF;
END_IF;
{endregion}

// === 🔑 §6 CYCLE DE VIE, R9 ET GUIDE OPERATEUR ===
{region "§6 Guide operateur & sorties"}
MachineHomingActive := HomingStarted;
Lifecycle.Busy      := HomingStarted;
Lifecycle.Done      := CommitPublished;

// Qualification de sortie — calcul UNIQUE, apres le deroule de transaction (§5) : un commit
// atomique OU un abandon du meme scan est immediatement reflete (comportement d'origine).
CommitOrOffsetValid := CommitPublished OR BucketOffsetValid;
MachineHomed := AxisHomed AND CommitOrOffsetValid
                AND NOT MachineHomingFailed AND NOT ReHomingAckRequired
                AND NOT Fault.Latched;

// R9 : capture de l'etape au front d'apparition du defaut latche, avant recalcul du guide.
IF LatchedEdge.Q THEN
    MachineHomingStepAtError := MachineHomingStep;
END_IF;

// Guide operateur — priorite decroissante, textes conserves a l'identique.
IF MachineHomingFailed THEN
    MachineHomingStep := E_MachineHomingStep.FAILED;
    MachineHomingInstruction := 'Referencement incomplet : rester en N2 et recommencer';
ELSIF MachineHomingLossSafeStop THEN
    MachineHomingStep := E_MachineHomingStep.LOSS_SAFESTOP;
    MachineHomingInstruction := 'Reference perdue en mouvement : arret controle en cours';
ELSIF HomingStarted OR M1Status.HomingBusy OR M2Status.HomingBusy THEN
    MachineHomingStep := E_MachineHomingStep.HOMING_IN_PROGRESS;
    MachineHomingInstruction := 'Referencement conjoint M1/M2 en cours : ne pas manoeuvrer';
ELSIF NOT M1Status.HomedAndReliable AND NOT M2Status.HomedAndReliable THEN
    MachineHomingStep := E_MachineHomingStep.BOTH_NOT_HOMED;
    MachineHomingInstruction := 'Codeurs M1 et M2 non references : passer en maintenance N2';
ELSIF NOT M1Status.HomedAndReliable THEN
    MachineHomingStep := E_MachineHomingStep.M1_NOT_HOMED;
    MachineHomingInstruction := 'Codeur M1 non reference ou mesure douteuse : homer M1';
ELSIF NOT M2Status.HomedAndReliable THEN
    MachineHomingStep := E_MachineHomingStep.M2_NOT_HOMED;
    MachineHomingInstruction := 'Codeur M2 non reference ou mesure douteuse : homer M2';
ELSIF NOT (CommitPublished OR BucketOffsetValid) THEN
    IF Mode <> E_Mode.MAINT_N2 THEN
        MachineHomingStep := E_MachineHomingStep.OFFSET_UNKNOWN;
        MachineHomingInstruction := 'Offset benne inconnu : passer en maintenance N2';
    ELSIF NOT TopPositionActive THEN
        MachineHomingStep := E_MachineHomingStep.NEED_TOP_POSITION;
        MachineHomingInstruction := 'Monter Both a vitesse lente jusqu au capteur haut';
    ELSIF NOT WinchesMechanicallyStopped THEN
        MachineHomingStep := E_MachineHomingStep.NEED_MECHANICAL_STOP;
        MachineHomingInstruction := 'Capteur haut atteint : relacher la commande et attendre l arret';
    ELSE
        MachineHomingStep := E_MachineHomingStep.AWAIT_BUCKET_CONFIRM;
        MachineHomingInstruction := 'Confirmer visuellement la benne : Fermee ou Ouverte';
    END_IF;
ELSE
    MachineHomingStep := E_MachineHomingStep.VALID;
    MachineHomingInstruction := 'Referencement machine valide : mode nominal disponible';
END_IF;

Ready := Enable AND NOT Fault.Latched;
{endregion}

END_FUNCTION_BLOCK
